       // //ABSOLUTE ENCODER
       IF #VTD_Control.AE_Error > 0 THEN
           "Set_Bit_F"(Bit := 5,
                       Bit_Value := 1,
                       Var := #VTD_Control.VTD_Errors.Error_Word_3);
       END_IF;

       //Errors while running
       IF #VTD_Control.Running THEN
           IF NOT (#VTD_Control.LP_State = 2) AND
               (#VTD_Control.LE > (#VTD_Settings.Teach_Values.Levels_LE[#LevelBelowExtractor] + #VTD_Settings.Slowdown_Count_LE) AND #VTD_Control.Instruction.Manual_Down)
               OR
               #IEC_Timer_0_Instance.Q
           THEN //22:4
               "Set_Bit_F"(Bit := 11,
                           Bit_Value := 1,
                           Var := #VTD_Control.VTD_Errors.Error_Word_1);
           END_IF;

           IF #VTD_Control.VFD_Error > 0 THEN //25:1
               "Set_Bit_F"(Bit := 0,
                           Bit_Value := 1,
                           Var := #VTD_Control.VTD_Errors.Error_Word_4);
           ELSIF #VTD_Control.LE_Error > 0 THEN //25:2
               "Set_Bit_F"(Bit := 1,
                           Bit_Value := 1,
                           Var := #VTD_Control.VTD_Errors.Error_Word_4);
           ELSIF #VTD_Control.AE_Error > 0 THEN //25:3
               "Set_Bit_F"(Bit := 2,
                           Bit_Value := 1,
                           Var := #VTD_Control.VTD_Errors.Error_Word_4);
           ELSIF (#LPL_Extended AND #LPL_Retracted) OR (#LPR_Extended AND #LPR_Retracted) THEN // 25:4
               "Set_Bit_F"(Bit := 3,
                           Bit_Value := 1,
                           Var := #VTD_Control.VTD_Errors.Error_Word_4);
           ELSIF #Lower_Limit AND NOT #Upper_limit THEN // 25:5
               "Set_Bit_F"(Bit := 4,
                           Bit_Value := 1,
                           Var := #VTD_Control.VTD_Errors.Error_Word_4);
           ELSIF NOT #Lower_Limit AND #Upper_limit THEN // 25:6
               "Set_Bit_F"(Bit := 5,
                           Bit_Value := 1,
                           Var := #VTD_Control.VTD_Errors.Error_Word_4);
           ELSIF #Lower_Limit AND #Upper_limit THEN // 25:7
               "Set_Bit_F"(Bit := 6,
                           Bit_Value := 1,
                           Var := #VTD_Control.VTD_Errors.Error_Word_4);
           END_IF;
       END_IF;

       //Check if overtravel limit switches has been hit
       IF #Upper_limit AND #Ultimate_Slow AND #Ulitmate_Creep AND #VTD_Control.Instruction.Manual_Up
       THEN //24:6 Top overtravel limit reached.
           "Set_Bit_F"(Bit := 7,
                       Bit_Value := 1,
                       Var := #VTD_Control.VTD_Errors.Error_Word_2);
           IF #VTD_Control.Mode = 2 OR #VTD_Control.Mode = 3 THEN
               #State := 400;
           ELSE
               #State := 0;
           END_IF;
       ELSIF #Lower_Limit AND #Ultimate_Slow AND #Ulitmate_Creep AND #VTD_Control.Instruction.Manual_Down
       THEN //24:7 Bottom overtravel limit reached.
               #VTD_Control.Error := TRUE; 
               "Set_Bit_F"(Bit := 8,
                           Bit_Value := 1,
                           Var := #VTD_Control.VTD_Errors.Error_Word_2);
               IF #VTD_Control.Mode = 2 OR #VTD_Control.Mode = 3 THEN
                   #State := 400;
               ELSE
                   #State := 0;
               END_IF;
       // ELSIF #Lower_Limit AND #Ultimate_Slow AND #Ulitmate_Creep AND #VTD_Control.Mode <> 4 THEN
       //     #VTD_Control.Instruction.Stop := TRUE;
       //     #VTD_Control.Error := TRUE; //24:7 Bottom Overtravel limit reached.
       //     "Set_Bit_F"(Bit := 8,
       //                 Bit_Value := 1,
       //                 Var := #VTD_Control.VTD_Errors.Error_Word_2);
       //     IF #VTD_Control.Mode = 2 OR #VTD_Control.Mode = 3 THEN
       //         #State := 400;
       //     ELSE
       //         #State := 0;
       //     END_IF;
       END_IF;

       //Need to monitor both encoders to (Need to uncomment)
       // #VTD_Control.Encoder_Delta := (#VTD_Control.LE - ((#VTD_Control.AE * #VTD_Settings.AE_Ratio)) * #VTD_Settings.Encoder_Delta_W1) + (#VTD_Control.Encoder_Delta * #VTD_Settings.Encoder_Delta_W2);
       IF ABS(#VTD_Control.Encoder_Delta) > #VTD_Settings.Encoder_Delta_Warning THEN
           //Send warning message that encoder error is to large
           #VTD_Control.Warning := 0;
       END_IF;

       "IEC_Timer_0_DB_10".TON(IN:=ABS(#VTD_Control.Encoder_Delta) > #VTD_Settings.Encoder_Delta_Error,
                               PT:=t#500ms);

       IF "IEC_Timer_0_DB_10".Q THEN
           //Send error message that encoder error is to large
           #VTD_Control.Error := TRUE; // 24:1
           "Set_Bit_F"(Bit := 2,
                       Bit_Value := 1,
                       Var := #VTD_Control.VTD_Errors.Error_Word_2);
           #State := 400;
       END_IF;

       // Level detect timer 
       IF #LD_Timer.Q THEN
           #LD_Timer(IN := FALSE,
                     PT := T#0s);
           #VTD_Control.Error := TRUE; // 24:10 VTD not level
           "Set_Bit_F"(Bit := 11,
                       Bit_Value := 1,
                       Var := #VTD_Control.VTD_Errors.Error_Word_4);
           #State := 400;
       END_IF;

       //Locking pin timer
       IF #LP_Timer.Q AND (#LPL_Retract OR #LPL_Extend) THEN //24:2 Locking pins took to long to extend
           "Set_Bit_F"(Bit := 3,
                       Bit_Value := 1,
                       Var := #VTD_Control.VTD_Errors.Error_Word_2);
       ELSIF #LP_Timer.Q AND (#LPR_Retract AND #LPR_Extend) THEN //24:3 Locking pins took to long to retract
           "Set_Bit_F"(Bit := 4,
                       Bit_Value := 1,
                       Var := #VTD_Control.VTD_Errors.Error_Word_2);
       END_IF;

       IF #Interlock_Timer.Q THEN //Interlock process timed out
           "Set_Bit_F"(Bit := 3,
                       Bit_Value := 1,
                       Var := #VTD_Control.VTD_Errors.Error_Word_3);
           #I_State := 400;
       END_IF;

       // Watchdog bit
       IF #Watchdog.Q THEN
           #VTD_Control.Running := FALSE;
           IF #VTD_Control.Mode = 4 THEN //24:9 Teach timed out
               "Set_Bit_F"(Bit := 10,
                           Bit_Value := 1,
                           Var := #VTD_Control.VTD_Errors.Error_Word_2);
           ELSIF #VTD_Control.Mode = 3 THEN //24:9 Auto timed out
               "Set_Bit_F"(Bit := 10,
                           Bit_Value := 1,
                           Var := #VTD_Control.VTD_Errors.Error_Word_2);
           ELSIF #VTD_Control.Mode = 2 THEN //24:9 Semi auto timed out
               "Set_Bit_F"(Bit := 10,
                           Bit_Value := 1,
                           Var := #VTD_Control.VTD_Errors.Error_Word_2);
           END_IF;
       END_IF;

       // go to error state
       IF  #VTD_Control.VTD_Errors.Error_Word_1 <> 0 OR
           #VTD_Control.VTD_Errors.Error_Word_2 <> 0 OR
           #VTD_Control.VTD_Errors.Error_Word_3 <> 0 OR
           #VTD_Control.VTD_Errors.Error_Word_4 <> 0 THEN
           #VTD_Control.Error := TRUE;
           #State := 400;
       END_IF;
   END_REGION

   REGION VFD
       //Status
       #VTD_Control.Motor.Ready := #SinaSpeed.Status = 16#7002;
       #VTD_Control.Motor.Running := #SinaSpeed.AxisEnabled;
       #VTD_Control.Motor.Error := #SinaSpeed.Status > 16#8000;

       //SETPOINT
       IF #VTD_Control.Motor_UP THEN
           #MainSetpoint := SCALE_X(MIN := 0,
                                    VALUE := NORM_X(MIN := 0,
                                                    VALUE := #VTD_Control.Motor_Speed,
                                                    MAX := 100),
                                    MAX := 1774);
       ELSIF #VTD_Control.Motor_Down THEN
           #MainSetpoint := (SCALE_X(MIN := 0,
                                     VALUE := NORM_X(MIN := 0,
                                                     VALUE := #VTD_Control.Motor_Speed,
                                                     MAX := 100),
                                     MAX := 1774)) * -1;
       ELSE
           #MainSetpoint := 0;
       END_IF;

       "IEC_Timer_0_DB".TON(IN:=#MainSetpoint <> 0,
                            PT:=T#500ms);

       IF "IEC_Timer_0_DB".Q THEN
           #MainSetpoint1 := #MainSetpoint;
       ELSE
           #MainSetpoint1 := 0;
       END_IF;

       IF #VTD_Control.Instruction.Enable THEN
           #SinaSpeed(EnableAxis := #VTD_Control.Motor_UP OR #VTD_Control.Motor_Down,
                          AckError := #VTD_Control.Instruction.Reset,
                          SpeedSp := #MainSetpoint1,
                          RefSpeed := 1774,
                          HWIDSTW := "VTD~PROFINET_interface~Standard_telegram_1",
                          HWIDZSW := "VTD~PROFINET_interface~Standard_telegram_1",
                          AxisEnabled => #VTD_Control.Motor.Status.%X0,
                          Lockout => #VTD_Control.Motor.Error,
                          Error => #VTD_Control.Motor.Error);
       END_IF;

       REGION Actual Speed
           IF #MainSetpoint1 > 0 THEN
               #VTD_Control.Motor.Speed_Actual := SCALE_X(MIN := 0,
                                                          VALUE := NORM_X(MIN := 0,
                                                                          VALUE := #SinaSpeed.ActVelocity,
                                                                          MAX := 1774),
                                                          MAX := 100);
           ELSIF #MainSetpoint1 < 0 THEN
               #VTD_Control.Motor.Speed_Actual := SCALE_X(MIN := 0,
                                                          VALUE := NORM_X(MIN := 0,
                                                                          VALUE := #SinaSpeed.ActVelocity * -1,
                                                                          MAX := 1774),
                                                          MAX := 100);
           ELSE
               #VTD_Control.Motor.Speed_Actual := 0;
           END_IF;
       END_REGION
   END_REGION

   //Assign local vars to outputs
   "Left LockingPin CMD Retract" := #LPL_Retract;
   "Left LockingPin CMD Extend" := #LPL_Extend;
   "Right LockingPin CMD Retract" := #LPR_Retract;
   "Right LockingPin CMD Extend" := #LPR_Extend;
END_FUNCTION_BLOCK

FUNCTION_BLOCK "EConveyor_FB"   // FB12, SCL
TITLE = Conveyor Instance FB
{ S7_Optimized_Access := 'TRUE' }
AUTHOR : Mertin Coetzee
VERSION : 0.1
// stored: AutoNumber true, IsIECCheckEnabled false, IsRetainMemResEnabled false, MemoryReserve 100, SetENOAutomatically false, UDAEnableTagReadback false
   VAR_INPUT
      Cnv_Settings : "ECnv_Settings";
      Cnv_Inputs : "ECnv_Inputs";
      VTD_Level : UInt;
      Cnv_TIP : Bool;
   END_VAR
   VAR_IN_OUT
      Cnv_Control : "ECnv_Control";
      SinaSpeed : SinaSpeed;
   END_VAR
   VAR
      State : UInt;
      Timer_TC : TON_TIME;
      Timer_Transfer { S7_SetPoint := 'True'} : TON_TIME;
      Watchdog { S7_SetPoint := 'True'} : TON_TIME;
      Transfer_Direction { S7_SetPoint := 'True'} : String;
      MainSetpoint : Int;
      SinaSpeed_Instance { S7_SetPoint := 'True'} : SinaSpeed;
      IEC_Timer_0_Instance_1 { S7_SetPoint := 'True'} : TON_TIME;
      IEC_Timer_0_Instance_2 { S7_SetPoint := 'True'} : TON_TIME;
      R_TRIG_Instance { S7_SetPoint := 'True'} : R_TRIG;
   END_VAR
   VAR_TEMP
      Execute_Old : Bool;
      Stop_Old : Bool;
      i : Int;
   END_VAR
BEGIN
   "R_TRIG_DB_15"(CLK := #Cnv_Control.Instruction.Execute AND NOT #Execute_Old);
   "R_TRIG_DB_16"(CLK := #Cnv_Control.Instruction.Stop AND NOT #Stop_Old);

   #Execute_Old := #Cnv_Control.Instruction.Execute;
   #Stop_Old := #Cnv_Control.Instruction.Stop;

   #Cnv_Control.Enabled := #Cnv_Control.Instruction.Enable;

   //MODES
   #Cnv_Control.Mode := #Cnv_Control.Instruction.Mode_Change;
   IF (#Cnv_Control.Mode = 1 OR #Cnv_Control.Mode = 5) AND NOT #Cnv_Control.Error THEN
       #State := 500;
   END_IF;

   #R_TRIG_Instance(CLK:=#Cnv_Control.Mode = 3);
   IF #R_TRIG_Instance.Q THEN
       #State := 0;
   END_IF;

   (*
   TODO:
   01. Need to add statemachine watchdog - Done
   02. Extractor needs to be on same floor for pallet to be moved in manual passed Rbwd - Done
   03. Complete reset state - Done
   04. Add stop inputs - Done
   05. Need to add variable motor speed, manual needs to be slower. - Done
   06. Need to add cyclic error checking. For odd sensor combinations as well - Partially done
   07. Need to add Shuttle monitor - Done
   08. Need to add Task ID check and start bit check to outbound pallet move. Check direction of pallet movement based on connected Cnv.
   09. Need to add checks for wrong direction of travel - Done
   10. Add checks for unsafe conditions with Cnv_Inputs - Partially Done
   11. Define Error codes - DOne
   12. Add watchdof time to Cnv Settings - Done
   13. Add self-timeout on manual 
   14. For shuttle in place sensor checks take into account extractor floor and safety stopper state
   15. Confirm modes and states are correct (Semi-auto and maintenance as well)
   16. Add the correct transfer process for the logistex-spacemaker pallet handovers.

   Mode select is done via the HMI. Might add external mode select switches.

           Mode select mask:
           0: Disabled
           1: Manual
           2: Semi-Auto
           3: Auto
           4: Teach - N/A for Cnv
           5: Maintenance

   Device ID Format: XXYYZZ    
   XX = Device type   
       01   VTD
       10  Cnv_Front_of_VTD
       11  Cnv_Rear_of_VTD
       12  Cnv_On_Extractor
       20  Safety_Stop_Front_of_VTD
       21  Safety_Stop_Rear_of_VTD
   YY = Floor   
   ZZ = VTD Connected to    
   Example: 110203 Conveyor at the rear of VTD 3 on level 2


    Sensor order for the conveyor:
    Lfwd Lpd1 Lpd2
     []   []   []
    ##############################
    #        Pallet Flow         #
    #         ------->>          #
    #                            #
    #                            #
    ##############################
                     []   []   []
                    Rpd2 Rpd1 Rbwd      
   *)

   REGION Cyclic Checks 
       #Cnv_Control.Cnv_Occupied := "Pallet in Position Rear VTD" AND "Pallet in Position Front VTD";

       //Check if a shuttle is in the Cnv
       FOR #i := 1 TO 3 DO
           IF "Shuttle_MQTT_DB".Shuttle_MQTT[#i].Message.Shuttle_Status.Position_ID = #Cnv_Settings.Barcode_ID THEN
               IF #Cnv_Inputs.Sdetect1 AND #Cnv_Inputs.Sdetect2 THEN
                   #Cnv_Control.Shuttle_In_Place := TRUE;
               ELSE
                   #Cnv_Control.Shuttle_In_Place := FALSE;
               END_IF;
           END_IF;
       END_FOR;

       // Update the Cnv_Control opbject
       #Cnv_Control.SM_State := #State;
       IF #Cnv_Control.Instruction.Inbound_Ready OR #Cnv_Control.Instruction.Outbound_Ready THEN
           #Cnv_Control.Ready_For_Task := TRUE;
       ELSE
           #Cnv_Control.Ready_For_Task := FALSE;
       END_IF;

   END_REGION

   REGION Auto/Semi/Manual mode
       CASE #State OF
           0: //IDLE MODE
               #Cnv_Control.Instruction.Transfer_Complete := 0;
               #Cnv_Control.Instruction.Transfer_in_Progress := FALSE;
               #Cnv_Control.Running := FALSE;
               #Cnv_Control.Motor.Forward := FALSE;
               #Cnv_Control.Motor.Reverse := FALSE;
               #Cnv_Control.Motor.Speed := 0;
               #Timer_Transfer(IN := FALSE,
                               PT := T#0S);
               IF #Cnv_Control.Enabled AND (#Cnv_Control.Mode = 3 OR #Cnv_Control.Mode = 2) AND #Cnv_Control.Error = 0 THEN
                   #State := 10;
               END_IF;

           10: //Standby - Conveyor ready to receive instruction
               IF ("R_TRIG_DB_15".Q OR #Cnv_Control.Instruction.Start_Transfer) AND "Control_DB".VTD_Control.Current_Level = #Cnv_Settings.Cnv_Level THEN
                   //Inbound Transfer
                   IF #Cnv_Control.Instruction.Inbound_Ready AND NOT #Cnv_Control.Running AND #Cnv_Control.Error = 0 AND
                       ("Control_DB".VTD_Control.Current_Level > 0 OR "Control_DB".PopUp_Cnv[2].Inputs."Lift Down")
                   THEN
                       #Cnv_Control.Done := FALSE;
                           #Cnv_Control.Running := TRUE;
                           #Cnv_Control.Instruction.Transfer_in_Progress := TRUE;
                           #Cnv_Control.Current_Task_ID := #Cnv_Control.Instruction.Task_ID;
                           #State := 20;

                       //Outbound Transfer    
                       ELSIF #Cnv_Control.Instruction.Outbound_Ready AND NOT #Cnv_Control.Running AND #Cnv_Control.Error = 0 AND
                           ("Control_DB".VTD_Control.Current_Level > 0 OR "Control_DB".PopUp_Cnv[2].Inputs."Lift Down")
                       THEN
                           #Cnv_Control.Done := FALSE;
                           #Cnv_Control.Running := TRUE;
                           #Cnv_Control.Instruction.Transfer_in_Progress := TRUE;
                           #Cnv_Control.Current_Task_ID := #Cnv_Control.Instruction.Task_ID;
                           #State := 30;
                   ELSE
                       #Cnv_Control.Warning := 1;// No task that can be started, yet start bit has been made true.
                   END_IF;
               ELSIF #Cnv_Control.Instruction.Start_Transfer AND "Control_DB".VTD_Control.Current_Level <> #Cnv_Settings.Cnv_Level THEN
                   //Extracot not at the correct level
                   "Set_Bit_F"(Bit := 2,
                               Bit_Value := 1,
                               Var := #Cnv_Control.Cnv_Errors.Error_Word_3);
               END_IF;

               //----------------------- Pallet Movement Inbound -----------------------
           20: // Running Roller FOWARD
               #Cnv_Control.Running := TRUE;
               #Cnv_Control.Motor.Forward := TRUE;
               #Cnv_Control.Motor.Speed := #Cnv_Settings.Full_Speed;
               #Transfer_Direction := 'Foward';

               IF "R_TRIG_DB_16".Q OR #Cnv_Control.Cnv_Occupied THEN
                   #Cnv_Control.Done := TRUE;
                   #Cnv_Control.Motor.Speed := 0;
                   #Cnv_Control.Motor.Forward := FALSE;
                   #Cnv_Control.Running := FALSE;
                   #State := 0;
               END_IF;

               //Monitor the transfer progress
               #Timer_Transfer(IN := TRUE,
                               PT := UINT_TO_TIME(#Cnv_Settings.Transfer_Time) * 1000);
               //If the watchdog bites, kill the process
               IF #Timer_Transfer.Q THEN //14:1 Transfer timed out
                   "Set_Bit_F"(Bit := 3,
                               Bit_Value := 1,
                               Var := #Cnv_Control.Cnv_Errors.Error_Word_2);
               END_IF;

               //----------------------- Pallet Movement Outbound -----------------------
           30: // Running Roller REVERSE
               IF (#VTD_Level = 0 AND "Control_DB".PopUp_Cnv[2].Chain_Motor.Status.%X0) OR
                   (#VTD_Level = 1 AND "Control_DB".LCnv_Control[1].Motor.Status.%X0) OR
                   (#VTD_Level = 2 AND "Control_DB".LCnv_Control[2].Motor.Status.%X0) OR
                   (#VTD_Level = 3 AND "Control_DB".LCnv_Control[3].Motor.Status.%X0) THEN
                   #Cnv_Control.Running := TRUE;
                   #Cnv_Control.Motor.Reverse := TRUE;
                   #Cnv_Control.Motor.Speed := #Cnv_Settings.Full_Speed;
                   #Transfer_Direction := 'Foward';
               END_IF;

               IF ("R_TRIG_DB_16".Q AND #Cnv_Control.Mode = 2) OR
                   (
                   (#VTD_Level = 0 AND NOT "PopUp Conveyor 2 - Pallet present 5") OR
                   (#VTD_Level = 1 AND NOT "Control_DB".LCnv_Control[1].Inputs."Pallet Detect 3") OR
                   (#VTD_Level = 2 AND NOT "Control_DB".LCnv_Control[2].Inputs."Pallet Detect 3") OR
                   (#VTD_Level = 3 AND NOT "Control_DB".LCnv_Control[3].Inputs."Pallet Detect 3") OR
                   (#VTD_Level = 99)
                   ) THEN
                   #Cnv_Control.Done := TRUE;
                   #Cnv_Control.Motor.Speed := 0;
                   #Cnv_Control.Motor.Forward := FALSE;
                   #Cnv_Control.Running := FALSE;
                   #State := 0;
               END_IF;

               //Monitor the transfer progress
               #Timer_Transfer(IN := TRUE,
                               PT := UINT_TO_TIME(#Cnv_Settings.Transfer_Time) * 1000);
               //If the watchdog bites, kill the process
               IF #Timer_Transfer.Q THEN //14:1 Transfer timed out
                   "Set_Bit_F"(Bit := 3,
                               Bit_Value := 1,
                               Var := #Cnv_Control.Cnv_Errors.Error_Word_2);
               END_IF;

           400: //Error state
               #Cnv_Control.Running := FALSE;
               #Cnv_Control.Motor.Speed := 0;
               #Cnv_Control.Motor.Forward := FALSE;
               #Cnv_Control.Motor.Reverse := FALSE;
               #Cnv_Control.Stopped := TRUE;
               #Cnv_Control.Instruction.Transfer_in_Progress := FALSE;
               #Watchdog(IN := FALSE,
                               PT := T#0S);
               #Timer_TC(IN := FALSE,
                               PT := T#0S);
               #Timer_Transfer(IN := FALSE,
                               PT := T#0S);
               #IEC_Timer_0_Instance_1(IN := FALSE,
                                       PT := T#0S);
               #IEC_Timer_0_Instance_2(IN := FALSE,
                                       PT := T#0S);
               IF #Cnv_Control.Instruction.Reset THEN
                   #Cnv_Control.Warning := 0;
                   #Cnv_Control.Current_Task_ID := 0;
                   #Cnv_Control.Error := FALSE; //Reset the conveyor

                   #Cnv_Control.Cnv_Errors.Error_Word_1 := 0;
                   #Cnv_Control.Cnv_Errors.Error_Word_2 := 0;
                   #Cnv_Control.Cnv_Errors.Error_Word_3 := 0;
                   #Cnv_Control.Cnv_Errors.Error_Word_4 := 0;
                   #State := 0;
               END_IF;

           500:
               IF #Cnv_Control.Enabled THEN
                   IF #"VTD_Level" = #Cnv_Settings.Cnv_Level THEN
                       IF #Cnv_Control.Instruction.Foward OR #Cnv_Control.Instruction.Start_Transfer THEN
                           #Cnv_Control.Motor.Speed := #Cnv_Settings.Manual_Speed;
                           #Cnv_Control.Motor.Forward := TRUE;
                           #Cnv_Control.Running := TRUE;
                       ELSIF #Cnv_Control.Instruction.Backward OR #Cnv_Control.Instruction.Start_Transfer_Backward THEN
                           #Cnv_Control.Motor.Speed := #Cnv_Settings.Manual_Speed;
                           #Cnv_Control.Motor.Reverse := TRUE;
                           #Cnv_Control.Running := TRUE;
                       ELSE
                           #Cnv_Control.Motor.Speed := 0;
                           #Cnv_Control.Motor.Forward := FALSE;
                           #Cnv_Control.Motor.Reverse := FALSE;
                           #Cnv_Control.Running := FALSE;
                       END_IF;
                   END_IF;
               END_IF;
               IF #Cnv_Control.Mode <> 1 AND #Cnv_Control.Mode <> 5 THEN
                   #State := 0;
               END_IF;
       END_CASE;
   END_REGION


   REGION Cyclic Error Checks
       IF NOT "Main_Safety_RTG1_DB".SAFETY_OK_VTD THEN //21:1
           "Set_Bit_F"(Bit := 0,
                       Bit_Value := 1,
                       Var := #Cnv_Control.Cnv_Errors.Error_Word_1);
       END_IF;

       IF #Cnv_Control.Motor.Error THEN
           "Set_Bit_F"(Bit := 0,
                       Bit_Value := 1,
                       Var := #Cnv_Control.Cnv_Errors.Error_Word_4);
       END_IF;


       // Shuttle in Place Cnv_Inputs - Need to confirm the order of these Cnv_Inputs.
       // IF (#Cnv_Settings.ID > 110000 AND #Cnv_Settings.ID < 120000 AND NOT #Cnv_Control.Inputs.Sdetect1 AND #Cnv_Control.Inputs.Sdetect2)
       //     OR (#Cnv_Settings.ID > 120000 AND #Cnv_Settings.ID < 130000 AND NOT #Cnv_Control.Inputs.Sdetect1 AND #Cnv_Control.Inputs.Sdetect2)
       // THEN //14:5 Shuttle is about to yeet itself down the VTD shaft
       //     "Set_Bit_F"(Bit := 7,
       //                 Bit_Value := 1,
       //                 Var := #Cnv_Control.Cnv_Errors.Error_Word_2);
       // END_IF;

       // IF (#Cnv_Settings.ID > 110000 AND #Cnv_Settings.ID < 120000 AND #Cnv_Control.Inputs.Sdetect1 AND NOT #Cnv_Control.Inputs.Sdetect2)
       //     OR (#Cnv_Settings.ID > 120000 AND #Cnv_Settings.ID < 130000 AND #Cnv_Control.Inputs.Sdetect1 AND NOT #Cnv_Control.Inputs.Sdetect2) THEN
       //     #Cnv_Control.Warning := 1; //Shuttle detected in conveyor not yet on barcode
       // END_IF;

       //Watchdog auto starts the moment any form of transfer occurs.
       // IF #State > 10 AND #State < 400 THEN
       //     #Watchdog(IN := TRUE,
       //               PT := T#600s);
       // ELSE
       //     #Watchdog.IN := FALSE;
       // END_IF;

       // IF #Watchdog.Q THEN
       //     #Watchdog.IN := FALSE;
       //     #Cnv_Control.Error := TRUE; //14:2  Watchdog bit
       //     "Set_Bit_F"(Bit := 4,
       //                 Bit_Value := 1,
       //                 Var := #Cnv_Control.Cnv_Errors.Error_Word_2);
       //     #State := 400;
       // END_IF;

       // go to error state
       IF #Cnv_Control.Cnv_Errors.Error_Word_1 <> 0 OR
           #Cnv_Control.Cnv_Errors.Error_Word_2 <> 0 OR
           #Cnv_Control.Cnv_Errors.Error_Word_3 <> 0 OR
           #Cnv_Control.Cnv_Errors.Error_Word_4 <> 0
           THEN
               #Cnv_Control.Error := TRUE;
               #State := 400;
       END_IF;
   END_REGION

   REGION VFD
       //Status
       #Cnv_Control.Motor.Ready := NOT #Cnv_Control.Motor.Error;

       #SinaSpeed(EnableAxis := #Cnv_Control.Motor.Forward OR #Cnv_Control.Motor.Reverse,
                  AckError := #Cnv_Control.Instruction.Reset,
                  SpeedSp := #MainSetpoint,
                  RefSpeed := 1745.0,
                  HWIDSTW := #Cnv_Settings.G120_Hardware_ID,
                  HWIDZSW := #Cnv_Settings.G120_Hardware_ID,
                  AxisEnabled => #Cnv_Control.Motor.Status.%X0,
                  Lockout => #Cnv_Control.Motor.Error,
                  Error => #Cnv_Control.Motor.Error);

       //MAIN SETPOINT
       IF #Cnv_Control.Motor.Reverse THEN
           #MainSetpoint := (SCALE_X(MIN := 0,
                                    VALUE := NORM_X(MIN := 0,
                                                    VALUE := #Cnv_Control.Motor.Speed,
                                                    MAX := 100),
                                    MAX := 1745.0)) * -1;
      ELSIF #Cnv_Control.Motor.Forward THEN
           #MainSetpoint := SCALE_X(MIN := 0,
                                     VALUE := NORM_X(MIN := 0,
                                                     VALUE := #Cnv_Control.Motor.Speed,
                                                     MAX := 100),
                                     MAX := 1745.0);
       ELSE
           #MainSetpoint := 0;
       END_IF;

       //Actual Speed
       IF #MainSetpoint > 0 THEN
           #Cnv_Control.Motor.Speed_Actual := SCALE_X(MIN := 0,
                                                      VALUE := NORM_X(MIN := 0,
                                                                      VALUE := #SinaSpeed.ActVelocity,
                                                                      MAX := 1745.0),
                                                      MAX := 100);
       ELSIF #MainSetpoint < 0 THEN
           #Cnv_Control.Motor.Speed_Actual := SCALE_X(MIN := 0,
                                                      VALUE := NORM_X(MIN := 0,
                                                                      VALUE := #SinaSpeed.ActVelocity * -1,
                                                                      MAX := 1745.0),
                                                      MAX := 100);
       ELSE
           #Cnv_Control.Motor.Speed_Actual := 0;
       END_IF;
   END_REGION
END_FUNCTION_BLOCK

FUNCTION_BLOCK "Buffer_Conveyor_FB"   // FB5, SCL
TITLE = Conveyor Instance FB
{ S7_Optimized_Access := 'TRUE' }
AUTHOR : Mertin Coetzee
VERSION : 0.1
// stored: AutoNumber true, IsIECCheckEnabled false, IsRetainMemResEnabled false, MemoryReserve 100, SetENOAutomatically false, UDAEnableTagReadback false
   VAR_INPUT
      Cnv_Settings : "Buffer_Cnv_Settings";
      VTD_Level : UInt;
      ECnv_TIP : Bool;
   END_VAR
   VAR_IN_OUT
      Cnv_Control : "Buffer_Cnv_Control";
      SinaSpeed : SinaSpeed;
   END_VAR
   VAR
      State : UInt;
      Timer_TC : TON_TIME;
      Timer_Transfer { S7_SetPoint := 'True'} : TON_TIME;
      Watchdog { S7_SetPoint := 'True'} : TON_TIME;
      Transfer_Direction { S7_SetPoint := 'True'} : String;
      MainSetpoint : Int;
      IEC_Timer_0_Instance_1 { S7_SetPoint := 'True'} : TON_TIME;
      R_TRIG_Instance { S7_SetPoint := 'True'} : R_TRIG;
   END_VAR
   VAR_TEMP
      Execute_Old : Bool;
      Stop_Old : Bool;
   END_VAR
BEGIN
   "R_TRIG_DB_17"(CLK := #Cnv_Control.Instruction.Execute AND NOT #Execute_Old);
   "R_TRIG_DB_18"(CLK := #Cnv_Control.Instruction.Stop AND NOT #Stop_Old);

   #Execute_Old := #Cnv_Control.Instruction.Execute;
   #Stop_Old := #Cnv_Control.Instruction.Stop;

   #Cnv_Control.Enabled := #Cnv_Control.Instruction.Enable;

   //MODES
   #Cnv_Control.Mode := #Cnv_Control.Instruction.Mode_Change;
   IF (#Cnv_Control.Mode = 1 OR #Cnv_Control.Mode = 5) AND NOT #Cnv_Control.Error THEN
       #State := 500;
   END_IF;

   #R_TRIG_Instance(CLK:=#Cnv_Control.Mode = 3);
   IF #R_TRIG_Instance.Q THEN
       #State := 0;
   END_IF;

   (*
   TODO:
   01. Need to add statemachine watchdog - Done
   02. Extractor needs to be on same floor for pallet to be moved in manual passed Rbwd - Done
   03. Complete reset state - Done
   04. Add stop inputs - Done
   05. Need to add variable motor speed, manual needs to be slower. - Done
   06. Need to add cyclic error checking. For odd sensor combinations as well - Partially done
   07. Need to add Shuttle monitor - Done
   08. Need to add Task ID check and start bit check to outbound pallet move. Check direction of pallet movement based on connected Cnv.
   09. Need to add checks for wrong direction of travel - Done
   10. Add checks for unsafe conditions with Cnv_Inputs - Partially Done
   11. Define Error codes - DOne
   12. Add watchdof time to Cnv Settings - Done
   13. Add self-timeout on manual 
   14. For shuttle in place sensor checks take into account extractor floor and safety stopper state
   15. Confirm modes and states are correct (Semi-auto and maintenance as well)
   16. Add the correct transfer process for the logistex-spacemaker pallet handovers.

   Mode select is done via the HMI. Might add external mode select switches.

           Mode select mask:
           0: Disabled
           1: Manual
           2: Semi-Auto
           3: Auto
           4: Teach - N/A for Cnv
           5: Maintenance

   Device ID Format: XXYYZZ    
   XX = Device type   
       40  VTD
       10  Cnv_Front_of_VTD
       11  Cnv_Rear_of_VTD
       12  Cnv_On_Extractor
       20  Safety_Stop_Front_of_VTD
       21  Safety_Stop_Rear_of_VTD

   YY = Floor   
   ZZ = VTD Connected to    
   Example: 110203 Conveyor at the rear of VTD 3 on level 2

   Pallet Alignment
   0 = no alignment
   1 = center alignment
   2 = Left
   3 = Right

    Sensor order for the conveyor:
    Lfwd Lpd1 Lpd2
     []   []   []
    ##############################
    #        Pallet Flow         #
    #         ------->>          #
    #                            #
    #                            #
    ##############################
                     []   []   []
                    Rpd2 Rpd1 Rbwd      
   *)

   REGION Cyclic Checks    
       #Cnv_Control.Cnv_Occupied := NOT #Cnv_Control.Inputs."Pallet Detect 1" AND (*#Cnv_Control."Inputs"."Pallet Detect 2" AND*) NOT #Cnv_Control.Inputs."Pallet Detect 3";

       //Check if a shuttle is in the Cnv
       IF NOT #Cnv_Control.Inputs.Sdetect1 AND NOT #Cnv_Control.Inputs.Sdetect2 THEN
           #Cnv_Control.Shuttle_In_Place := TRUE;
       ELSE
           #Cnv_Control.Shuttle_In_Place := FALSE;
       END_IF;

       // Update the Cnv_Control opbject
       #Cnv_Control.SM_State := #State;
       #Cnv_Control.Stopped := NOT #Cnv_Control.Running;
       IF #Cnv_Control.Instruction.Inbound_Ready OR #Cnv_Control.Instruction.Outbound_Ready THEN
           #Cnv_Control.Ready_For_Task := TRUE;
       ELSE
           #Cnv_Control.Ready_For_Task := FALSE;
       END_IF;

   END_REGION

   REGION Auto/Semi auto mode
       CASE #State OF
           0: //Initialization
               #Cnv_Control.Instruction.Transfer_Complete := 0;
               #Cnv_Control.Instruction.Transfer_in_Progress := FALSE;
               #Cnv_Control.Running := FALSE;
               #Cnv_Control.Motor.Forward := FALSE;
               #Cnv_Control.Motor.Reverse := FALSE;
               #Cnv_Control.Motor.Speed := 0;
               #Timer_Transfer(IN := FALSE,
                               PT := T#0S);
               IF #Cnv_Control.Enabled AND (#Cnv_Control.Mode = 3 OR #Cnv_Control.Mode = 2) AND #Cnv_Control.Error = 0 THEN
                   #State := 10;
               END_IF;

               10: //Standby - Conveyor ready to receive instruction
                   IF ("R_TRIG_DB_17".Q OR #Cnv_Control.Instruction.Start_Transfer) AND "Control_DB".VTD_Control.Current_Level = #Cnv_Settings.Cnv_Level THEN
                       //Inbound Transfer
                       IF #Cnv_Control.Instruction.Inbound_Ready AND NOT #Cnv_Control.Running AND #Cnv_Control.Error = 0 THEN
                           //Check transfer ID
                           #Cnv_Control.Done := FALSE;
                               #Cnv_Control.Running := TRUE;
                               #Cnv_Control.Instruction.Transfer_in_Progress := TRUE;
                               #Cnv_Control.Current_Task_ID := #Cnv_Control.Instruction.Task_ID;
                               #State := 20;

                           //Outbound Transfer    
                       ELSIF #Cnv_Control.Instruction.Outbound_Ready AND NOT #Cnv_Control.Running AND #Cnv_Control.Error = 0 THEN
                           //Check transfer ID
                           #Cnv_Control.Done := FALSE;
                               #Cnv_Control.Running := TRUE;
                               #Cnv_Control.Instruction.Transfer_in_Progress := TRUE;
                               #Cnv_Control.Current_Task_ID := #Cnv_Control.Instruction.Task_ID;
                               #State := 30;
                       ELSE
                           #Cnv_Control.Warning := 0;// No task that can be started, yet start bit has been made true.
                       END_IF;
                   ELSIF #Cnv_Control.Instruction.Start_Transfer AND "Control_DB".VTD_Control.Current_Level <> #Cnv_Settings.Cnv_Level THEN
                       //Extractor not at the correct level
                       "Set_Bit_F"(Bit := 2,
                                   Bit_Value := 1,
                                   Var := #Cnv_Control.Cnv_Errors.Error_Word_3);
                   END_IF;

                   //----------------------- Pallet Movement Inbound -----------------------
               20: // Running Roller FOWARD
                   #Cnv_Control.Running := TRUE;
                   #Cnv_Control.Motor.Forward := TRUE;
                   #Cnv_Control.Motor.Speed := #Cnv_Settings.Full_Speed;
                   #Transfer_Direction := 'Foward';

                   IF "R_TRIG_DB_18".Q OR NOT #Cnv_Control.Inputs."Pallet Detect 3" THEN
                       #Cnv_Control.Done := TRUE;
                       #Cnv_Control.Motor.Speed := 0;
                       #Cnv_Control.Motor.Forward := FALSE;
                       #Cnv_Control.Running := FALSE;
                       #State := 0;
                   END_IF;

                   //Monitor the transfer progress
                   #Timer_Transfer(IN := TRUE,
                                   PT := UINT_TO_TIME(#Cnv_Settings.Transfer_Time) * 1000);
                   //If the watchdog bites, kill the process
                   IF #Timer_Transfer.Q THEN //14:1 Transfer timed out
                       "Set_Bit_F"(Bit := 3,
                                   Bit_Value := 1,
                                   Var := #Cnv_Control.Cnv_Errors.Error_Word_2);
                   END_IF;

                   //----------------------- Pallet Movement Outbound -----------------------
               30: // Running Roller REVERSE
                   #Cnv_Control.Running := TRUE;
                   #Cnv_Control.Motor.Reverse := TRUE;
                   #Cnv_Control.Motor.Speed := #Cnv_Settings.Full_Speed;
                   #Transfer_Direction := 'Foward';

                   IF "R_TRIG_DB_18".Q OR "Control_DB".ECnv_Control.Cnv_Occupied THEN
                       #Cnv_Control.Done := TRUE;
                       #Cnv_Control.Motor.Speed := 0;
                       #Cnv_Control.Motor.Forward := FALSE;
                       #Cnv_Control.Running := FALSE;
                       #State := 0;
                   END_IF;

                   //Monitor the transfer progress
                   #Timer_Transfer(IN := TRUE,
                                   PT := UINT_TO_TIME(#Cnv_Settings.Transfer_Time) * 1000);
                   //If the watchdog bites, kill the process
                   IF #Timer_Transfer.Q THEN //14:1 Transfer timed out
                       "Set_Bit_F"(Bit := 3,
                                   Bit_Value := 1,
                                   Var := #Cnv_Control.Cnv_Errors.Error_Word_2);
                   END_IF;

               400: //Error state
                   #Cnv_Control.Running := FALSE;
                   #Cnv_Control.Motor.Speed := 0;
                   #Cnv_Control.Motor.Forward := FALSE;
                   #Cnv_Control.Motor.Reverse := FALSE;
                   #Cnv_Control.Instruction.Stop := FALSE;
                   #Cnv_Control.Instruction.Transfer_in_Progress := FALSE;
                   #Watchdog(IN := FALSE,
                                   PT := T#0S);
                   #Timer_TC(IN := FALSE,
                                   PT := T#0S);
                   #Timer_Transfer(IN := FALSE,
                                   PT := T#0S);
                   #IEC_Timer_0_Instance_1(IN := FALSE,
                                           PT := T#0S);
                   IF #Cnv_Control.Instruction.Reset THEN
                       #Cnv_Control.Warning := 0;
                       #Cnv_Control.Current_Task_ID := 0;
                       #Cnv_Control.Error := FALSE; //Reset the conveyor

                       #Cnv_Control.Cnv_Errors.Error_Word_1 := 0;
                       #Cnv_Control.Cnv_Errors.Error_Word_2 := 0;
                       #Cnv_Control.Cnv_Errors.Error_Word_3 := 0;
                       #Cnv_Control.Cnv_Errors.Error_Word_4 := 0;
                       #State := 0;
                   END_IF;

               500:
                   IF #Cnv_Control.Enabled THEN
                       IF #Cnv_Control.Instruction.Foward OR #Cnv_Control.Instruction.Start_Transfer THEN
                               #Cnv_Control.Motor.Speed := #Cnv_Settings.Manual_Speed;
                               #Cnv_Control.Motor.Forward := TRUE;
                               #Cnv_Control.Running := TRUE;
                           ELSIF #Cnv_Control.Instruction.Backward OR #Cnv_Control.Instruction.Start_Transfer_Backward THEN
                               #Cnv_Control.Motor.Speed := #Cnv_Settings.Manual_Speed;
                               #Cnv_Control.Motor.Reverse := TRUE;
                               #Cnv_Control.Running := TRUE;
                           ELSE
                               #Cnv_Control.Motor.Speed := 0;
                               #Cnv_Control.Motor.Forward := FALSE;
                               #Cnv_Control.Motor.Reverse := FALSE;
                               #Cnv_Control.Running := FALSE;
                           END_IF;
                       END_IF;
                   IF #Cnv_Control.Mode <> 1 AND #Cnv_Control.Mode <> 5 THEN
                       #State := 0;
                   END_IF;
           END_CASE;
       END_REGION



   REGION Cyclic Error Checks
       IF NOT "Main_Safety_RTG1_DB".SAFETY_OK_VTD THEN //11:1
           "Set_Bit_F"(Bit := 0,
                       Bit_Value := 1,
                       Var := #Cnv_Control.Cnv_Errors.Error_Word_1);
       END_IF;

       // IF #Cnv_Control.Instruction.Stop THEN //11:2
       //     "Set_Bit_F"(Bit := 1,
       //                 Bit_Value := 1,
       //                 Var := #Cnv_Control.Cnv_Errors.Error_Word_1);
       // END_IF;

       IF #Cnv_Control.Motor.Error THEN
           "Set_Bit_F"(Bit := 0,
                       Bit_Value := 1,
                       Var := #Cnv_Control.Cnv_Errors.Error_Word_4);
       END_IF;

       // Pallet Sensor Checks
       // IF #Cnv_Control.Inputs.Lfwd AND #Cnv_Control.Inputs.Rbwd THEN
       //     #Cnv_Control.Error := TRUE; //15:2 Combination of Cnv_Inputs indicates issue in conveyor
       //     "Set_Bit_F"(Bit := 1,
       //                 Bit_Value := 1,
       //                 Var := #Cnv_Control.Cnv_Errors.Error_Word_4);
       //     #State := 400;
       // IF #Cnv_Control.Inputs.Lfwd AND #Cnv_Control.Inputs.Lpd1 AND #Cnv_Control.Inputs.Rpd1 THEN
       //     #Cnv_Control.Error := TRUE; //15:3 Combination of Cnv_Inputs indicates issue in conveyor
       //     "Set_Bit_F"(Bit := 2,
       //                 Bit_Value := 1,
       //                 Var := #Cnv_Control.Cnv_Errors.Error_Word_4);
       //     #State := 400;
       // ELSIF #Cnv_Control.Inputs.Rbwd AND #Cnv_Control.Inputs.Lpd1 AND #Cnv_Control.Inputs.Rpd1 THEN
       //     #Cnv_Control.Error := TRUE; //15:4 Combination of Cnv_Inputs indicates issue in conveyor
       //     "Set_Bit_F"(Bit := 3,
       //                 Bit_Value := 1,
       //                 Var := #Cnv_Control.Cnv_Errors.Error_Word_4);
       //     #State := 400;
       // END_IF;

       // Shuttle in Place Cnv_Inputs - Need to confirm the order of these Cnv_Inputs.
       // IF (#Cnv_Settings.ID > 110000 AND #Cnv_Settings.ID < 120000 AND NOT #Cnv_Control.Inputs.Sdetect1 AND #Cnv_Control.Inputs.Sdetect2)
       //     OR (#Cnv_Settings.ID > 120000 AND #Cnv_Settings.ID < 130000 AND NOT #Cnv_Control.Inputs.Sdetect1 AND #Cnv_Control.Inputs.Sdetect2) THEN
       //     #Cnv_Control.Error := TRUE; //14:5 Shuttle is about to yeet itself down the VTD shaft
       //     "Set_Bit_F"(Bit := 7,
       //                 Bit_Value := 1,
       //                 Var := #Cnv_Control.Cnv_Errors.Error_Word_2);
       //     #State := 400;
       // END_IF;

       // IF (#Cnv_Settings.ID > 110000 AND #Cnv_Settings.ID < 120000 AND #Cnv_Control.Inputs.Sdetect1 AND NOT #Cnv_Control.Inputs.Sdetect2)
       //     OR (#Cnv_Settings.ID > 120000 AND #Cnv_Settings.ID < 130000 AND #Cnv_Control.Inputs.Sdetect1 AND NOT #Cnv_Control.Inputs.Sdetect2) THEN
       //     #Cnv_Control.Warning := 0; //Shuttle detected in conveyor not yet on barcode
       // END_IF;

       // // #Watchdog auto starts the moment Any form OF transfer occurs.
       // IF #State > 10 AND #State < 400 THEN
       //     #Watchdog(IN := TRUE,
       //               PT := T#200s);
       // ELSE
       //     #Watchdog.IN := FALSE;
       // END_IF;

       // IF #Watchdog.Q THEN
       //     #Watchdog.IN := FALSE;
       //     #Cnv_Control.Error := TRUE; //14:2  Watchdog bit
       //     "Set_Bit_F"(Bit := 4,
       //                 Bit_Value := 1,
       //                 Var := #Cnv_Control.Cnv_Errors.Error_Word_2);
       //     #State := 400;
       // END_IF;

       // go to error state
       IF #Cnv_Control.Cnv_Errors.Error_Word_1 <> 0 OR
           #Cnv_Control.Cnv_Errors.Error_Word_2 <> 0 OR
           #Cnv_Control.Cnv_Errors.Error_Word_3 <> 0 OR
           #Cnv_Control.Cnv_Errors.Error_Word_4 <> 0
           THEN
               #Cnv_Control.Error := TRUE;
               #State := 400;
       END_IF;
   END_REGION

   REGION VFD
       //Status
       #Cnv_Control.Motor.Ready := NOT #Cnv_Control.Motor.Error;

       #SinaSpeed(EnableAxis := #Cnv_Control.Motor.Forward OR #Cnv_Control.Motor.Reverse,
                  AckError := #Cnv_Control.Instruction.Reset,
                  SpeedSp := #MainSetpoint,
                  RefSpeed := 1745.0,
                  HWIDSTW := #Cnv_Settings.G120_Hardware_ID,
                  HWIDZSW := #Cnv_Settings.G120_Hardware_ID,
                  AxisEnabled => #Cnv_Control.Motor.Status.%X0,
                  Lockout => #Cnv_Control.Motor.Error,
                  Error => #Cnv_Control.Motor.Error);

       //MAIN SETPOINT
       IF #Cnv_Control.Motor.Forward THEN
           #MainSetpoint := (SCALE_X(MIN := 0,
                                    VALUE := NORM_X(MIN := 0,
                                                    VALUE := #Cnv_Control.Motor.Speed * 1.681,
                                                    MAX := 100),
                                    MAX := 1745.0) * -1);
       ELSIF #Cnv_Control.Motor.Reverse THEN
           #MainSetpoint := SCALE_X(MIN := 0,
                                     VALUE := NORM_X(MIN := 0,
                                                     VALUE := #Cnv_Control.Motor.Speed * 1.681,
                                                     MAX := 100),
                                     MAX := 1745.0);
       ELSE
           #MainSetpoint := 0;
       END_IF;

       REGION Actual Speed
           IF #MainSetpoint > 0 THEN
               #Cnv_Control.Motor.Speed_Actual := SCALE_X(MIN := 0,
                                                          VALUE := NORM_X(MIN := 0,
                                                                          VALUE := #SinaSpeed.ActVelocity,
                                                                          MAX := 1745.0),
                                                          MAX := 100);
           ELSIF #MainSetpoint < 0 THEN
               #Cnv_Control.Motor.Speed_Actual := SCALE_X(MIN := 0,
                                                          VALUE := NORM_X(MIN := 0,
                                                                          VALUE := #SinaSpeed.ActVelocity * -1,
                                                                          MAX := 1745.0),
                                                          MAX := 100);
           ELSE
               #Cnv_Control.Motor.Speed_Actual := 0;
           END_IF;
       END_REGION
   END_REGION
END_FUNCTION_BLOCK

FUNCTION_BLOCK "Safety_Stops_FB"   // FB7, SCL
{ S7_Optimized_Access := 'TRUE' }
VERSION : 0.1
// stored: AutoNumber true, IsIECCheckEnabled false, IsRetainMemResEnabled false, MemoryReserve 100, SetENOAutomatically false, UDAEnableTagReadback false
   VAR_INPUT
      Mode : UInt;
      Timeout : UInt;
      Reset : Bool;
      Up : Bool;
      Down : Bool;
   END_VAR
   VAR_OUTPUT
      Rotate : Bool;
   END_VAR
   VAR_IN_OUT
      Sfts_Control : "Sfts_Control";
   END_VAR
   VAR
      State : UInt;
      LP_Timer { ExternalAccessible := 'False'; ExternalVisible := 'False'; ExternalWritable := 'False'} : TON_TIME;
      IEC_Timer_0_Instance { S7_SetPoint := 'True'} : TOF_TIME;
      Timer_1 : Time;
   END_VAR
BEGIN
   #Sfts_Control.Enabled := #Sfts_Control.Instruction.Enable := #Mode = 2 OR #Mode = 3;

   //MODES
   IF (#Mode = 1 OR #Mode = 5) AND NOT #Sfts_Control.Error THEN
       #State := 500;
   END_IF;

   (*
   TODO
   1. Need to add the mode and running checks for manual mode
   2. Add output for safety stop brake.

   Mode select is done via the HMI. Might add external mode select switches.

           Mode select mask:
           0: Disabled
           1: Manual
           2: Semi-Auto
           3: Auto
           4: Teach - N/A for Cnv
           5: Maintenance

   Device ID Format: XXYYZZ    
   XX = Device type   
       01   VTD
       10  Cnv_Front_of_VTD
       11  Cnv_Rear_of_VTD
       12  Cnv_On_Extractor
       20  Safety_Stop_Front_of_VTD
       21  Safety_Stop_Rear_of_VTD
   YY = Floor   
   ZZ = VTD Connected to 
   *)

   REGION Assign Inputs
       #Sfts_Control.Inputs.LP_Extended := #Up;
       #Sfts_Control.Inputs.LP_Retracted := #Down;
   END_REGION

   REGION Cyclic Checks
       //Update variables
       #Sfts_Control.SM_State := #State;

       #LP_Timer(IN := #Sfts_Control.Running,
                 PT := UINT_TO_TIME(#Timeout));

       //STOPPER STATE
       IF #Sfts_Control.Inputs.LP_Extended AND NOT #Sfts_Control.Inputs.LP_Retracted THEN
           #Sfts_Control.LP_State := 1; // EXTENDED
       ELSIF NOT #Sfts_Control.Inputs.LP_Extended AND #Sfts_Control.Inputs.LP_Retracted THEN
           #Sfts_Control.LP_State := 0; //RETRACTED
       ELSE
           #Sfts_Control.LP_State := 2; //LOST
       END_IF;;
   END_REGION

   REGION Auto Mode

           CASE #State OF
               0: //IDLE MODE
                   IF #Mode = 2 OR #Mode = 3 THEN
                       IF #Sfts_Control.Instruction.Enable AND #Sfts_Control.Error = 0 THEN
                           #Sfts_Control.Enabled := TRUE;
                           #State := 10;
                       END_IF;
                   END_IF;
               10: //Standby
                   IF NOT #Sfts_Control.Running AND #Sfts_Control.Error = 0 AND #Sfts_Control.Instruction.LP_Extend THEN
                       IF #Sfts_Control.Inputs.LP_Extended THEN
                           ; // Complete the task as the LP ar already extended
                       ELSIF #Sfts_Control.Inputs.LP_Retracted THEN
                           #Sfts_Control.Running := True;
                           #State := 20;
                       ELSE
                           #Sfts_Control.Error := 0; //Unknown locking pin state
                           #State := 400;
                       END_IF;
                   ELSIF NOT #Sfts_Control.Running AND #Sfts_Control.Error = 0 AND #Sfts_Control.Instruction.LP_Retract THEN
                       IF #Sfts_Control.Inputs.LP_Retracted THEN
                           ; // Complete the task as the LP ar already extended
                       ELSIF #Sfts_Control.Inputs.LP_Extended THEN
                           #Sfts_Control.Running := True;
                           #State := 40;
                       ELSE
                           #Sfts_Control.Error := 0; //Unknown locking pin state
                           #State := 400;
                       END_IF;
                   END_IF;

               20: //Extend safety locking pins
                   #Sfts_Control.Motor_Extend := TRUE;
                   IF #Sfts_Control.Inputs.LP_Extended THEN
                       #Sfts_Control.Motor_Extend := FALSE;
                       #Sfts_Control.Running := FALSE;
                       #State := 0;
                   END_IF;

               40: //Retract safety locking pins
                   #Sfts_Control.Motor_Retract := TRUE;
                   IF #Sfts_Control.Inputs.LP_Retracted THEN
                       #Sfts_Control.Motor_Retract := FALSE;
                       #Sfts_Control.Running := FALSE;
                       #State := 0;
                   END_IF;

               400: // Error#Sfts_Control
                   #Sfts_Control.Motor_Retract := FALSE;
                   #Sfts_Control.Motor_Extend := FALSE;
                   #Sfts_Control.Running := FALSE;
                   #LP_Timer(IN := FALSE,
                             PT := T#0S);
                   IF #Reset THEN
                       #Sfts_Control.Error := FALSE;
                       #State := 0;
                   END_IF;

               500:
                   IF #Sfts_Control.Instruction.Manual_Extend AND NOT #Sfts_Control.Inputs.LP_Extended THEN
                       #Sfts_Control.Motor_Extend := TRUE;
                       #Sfts_Control.Running := TRUE;
                   ELSIF #Sfts_Control.Instruction.Manual_Retract AND NOT #Sfts_Control.Inputs.LP_Retracted THEN
                       #Sfts_Control.Motor_Retract := TRUE;
                       #Sfts_Control.Running := TRUE;
                   ELSE
                       #Sfts_Control.Motor_Extend := FALSE;
                       #Sfts_Control.Motor_Retract := FALSE;
                       #Sfts_Control.Running := FALSE;
                   END_IF;

                   IF #Mode <> 1 AND #Mode <> 5 THEN
                       #State := 0;
                   END_IF;
           END_CASE;
   END_REGION

   REGION Cyclic Error Checks
       IF #Sfts_Control.Inputs.LP_Extended AND #Sfts_Control.Inputs.LP_Retracted THEN
           #Sfts_Control.Error := TRUE; //Cant have the locking pins extended and retracted at the same time11
       END_IF;

       // Statement section REGION
       IF #LP_Timer.Q THEN
           #Sfts_Control.Error := TRUE;//locking pin timeout
       END_IF;

       IF #Sfts_Control.Error THEN
           #State := 400;
       END_IF;
   END_REGION

   REGION Assign outputs
       #IEC_Timer_0_Instance(IN := #Sfts_Control.Motor_Extend OR #Sfts_Control.Motor_Retract,
                             PT := #Timer_1,
                             Q => #Rotate);
   END_REGION
END_FUNCTION_BLOCK

FUNCTION "Encoders" : Void   // FC8, SCL
{ S7_Optimized_Access := 'TRUE' }
VERSION : 0.1
// stored: AutoNumber true, IsIECCheckEnabled false, SetENOAutomatically false, UDAEnableTagReadback false
BEGIN
   REGION ABSOLUTE ENCODER
       //STATUS---------------------------------------------------------------------------------------------------------------------
       //
       //Encoder state word 2 - INPUT WORD 1
       //
       // 15 … 12 Encoder’s Sign-OF-Life (NOT relevant)
       // 11, 10 Reserved
       // 9 Control requested 0 = No control BY the PLC requested 1 = Control BY the PLC requested
       // 8 … 0 Reserved

       //Sensor 1 state word - INPUT WORD 2
       //
       // 15 Encoder error Description 0 = No error 1 = Error The error code is output in G1_XIST2.
       // 14 Park mode activated 0 = Normal operation 1 = Park mode activated Feedback based on G1_STW bit 14: No output OF position data G1_XIST1 AND G1_XIST2
       // 13 Transmission OF absolute position value 0 = No transmission 1 = Position value is output in G1_XIST2
       // 12 Status OF the Preset function (set/shift OF home position executed) 0 = No Preset function active 1 = Preset function is run Feedback based on G1_STW bit 12:  
       // 11 Requirement OF error acknowledgement detected New position value is output in G1_XIST1 AND G1_XIST2. On conclusion OF the Preset function the bit is set TO 0. 0 = No RETURN acknowledgement OF Encoder error 1 = Requirement OF error acknowledgement detected Reaction TO bit 15 in the sensor control word 1 G1_STW is acknowledged (see Table 14)
       // 10 Reserved
       // 9 … 0 NOT supported

       //Position 1 - INPUT WORD 3 AND 4
       // "AE_Position_1_Scaled" := (*SCALE_X(MIN := "Settings_DB".VTD_Settings.VTD_Min_Height,
       //                                   VALUE := *)NORM_X(MIN := 0,
       //                                                   VALUE := (SHL(IN:="AE_Position_1", N:=2) * 0.00228881) (*- "AE_Offset"*),
       //                                                   MAX := 1073741824)(*,
       //                                   MAX := "Settings_DB".VTD_Settings.VTD_Max_Heigh)*);
       // "mm_per_pulse" := 401,5584 / 262144;
       "AE_Position_1_Scaled" := (((1073741823 - (SHR(IN := "AE_Position_1", N := 2))) - 31381317) * 0.0015318237304688) - 1548572;
       // Position 2 - INPUT WORD 5 AND 6
       "AE_Position_2_Scaled" := SHR(IN := "AE_Position_2", N := 2);

       //Speed A - INPUT WORD 7
       "AE_Speed_Justified" := "AE_Speed";

       //CONTROL---------------------------------------------------------------------------------------------------------------------
       //
       //Encoder control word 2 - OUTPUT WORD 1
       //
       // 15 … 12 Master’s Sign-OF-Life (NOT relevant)
       // 10 control BY PLC 0 = No control BY the PLC 1 = Control BY the PLC Enables the PLC BY using control words TO activate / deactivate encoder functions
       // 7 Fault acknowledge Error-buffer handling NOT supported
       // 11, 9, 8, 6 … 0 Reserved
       // "AE_Control_Word_1".%X10 := "AE_PLC_Control";
       "AE_Control_Word_1".%X7 := "VTD_Reset_HMI_Tags";

       //Sensor 1 control word - OUTPUT WORD 2
       //
       // 15 Acknowledging a sensor error Description 0 = Encoder error message NOT acknowledged BY PLC 1 = Encoder error message acknowledged BY the PLC
       // 14 Activate park mode 0 = Normal operation 1 = Activate park mode
       // 13 Request FOR the absolute position value 0 = No request 1 = Request BY the master Results in the cyclic output OF the position values in G1_XIST2
       // 12 Activate preset value (see note below) Defines that a configured preset value is used (see section 3.5 on page 24) 0 = Preset value is NOT activated 1 = Preset value is activated
       // 11 Preset mode Defines how a configured preset value is used 0 = Preset value is used as a new absolute value 1 = Preset value is added TO the previous value
       // 10 … 0 Reserved
       // "AE_Control_Word_2".%X15 := "VTD_Reset_HMI_Tags";
       // "AE_Control_Word_2".%X14 := "AE_Activate_ParkMode";
       // "AE_Control_Word_2".%X13 := "AE_Request_ABS_Value";
       // "AE_Control_Word_2".%X12 := "AE_Activate_Preset_Value";
       // "AE_Control_Word_2".%X11 := "AE_Preset_Mode";
   END_REGION

   REGION LINEAR ENCODER
       "LE_X_Unsafe_Position_1" := DINT_TO_REAL("LE_X_Unsafe_Position") / 10;
       "LE_Speed_1" := "LE_Speed" * 10;
       //STATUS 
       //
       // 0 ERR - Error message (Error code in XP00– XP15); remaining bits = 0, see Error Codes
       // 1 NP - No position information/OUT (XP = 0, YP = 0, SP = 0)
       // 2 WRN - Warnings present, see Warning Module
       // 3 EV - Event present
       // 4 posdetected - Valid position information available

       //WARNINGS
       //
       // 0 WRN01 A code with non-PXV content was found.
       // 1 WRN02 the read head is too close TO the Data Matrix code tape.
       // 2 WRN03 the read head is too far from the Data Matrix code tape.
       // 3 WRN04 Y position too large. The sensor is just before OUT.
       // 4 WRN05 Y position is too small. The sensor is just before OUT.
       // 5 WRN06 the read head is rotated OR tilted in relation TO the Data Matrix code tape.
       // 6 WRN07 Low level OF code contrast.
       // 7 WRN08 Repair tape detected.
       // 8 WRN09 Temperature too high.
       // 9...15 Reserved

       //QUALITY GRADE
       //
       //The quality grades enable constant monitoring of the code tape and the camera along the entire
       //traverse distance. This enables you to detect and act upon potential damage or contamination
       //of the code tape and camera at the earliest stage possible during commissioning and normal
       //operation. As a result, this maximizes the overall functional reliability of your plant, and
       //it means you are able to immediately localize the issue in the case of a fault. Evaluations
       //are made using a scale of 1 to 6. The value 1 is the best possible read quality. A value greater
       //than 3 or worse requires the camera and its path to be inspected. The value 7 signifies "No position"
       //because no code was detected. An evaluation that indicates poor quality as the outcome can be due to
       //a misalignment or incorrect orientation, an incorrect measuring distance, or because the code tape has been affixed incorrectly
   END_REGION

       //RESET SAFETY POSITION LINEAR ENCODER
       "R_TRIG_DB_10"(CLK:="LE_Safe_Status" = 0);
       "Reintegration" := "R_TRIG_DB_10".Q;
END_FUNCTION

FUNCTION_BLOCK "FB_SICK_AFx60_PN"   // FB30, SCL
TITLE = SICK AFx60 PN
{ S7_Optimized_Access := 'TRUE' }
AUTHOR : SICKAG
FAMILY : SICKAG
VERSION : 1.1
// This function block simplifies the usage of the AFx60 encoder on Siemens S7-1200 /S7-1500 PLCs.
// It's support you to exchange the acyclic service data between the PLC and the AFx60 via Profinet (according to PROFIdrive V4.1).
// stored: AutoNumber true, IsIECCheckEnabled false, IsRetainMemResEnabled false, MemoryReserve 100, SetENOAutomatically false, UDAEnableTagReadback false
   VAR_INPUT
      ID : HW_IO;   // Hardware identifier of the "Parameter access point" module
      TOut : Time := T#5s;   // Timeout time
      Req : Bool;   // Positive trigger starts a request with the parameter set in the parameter selection
      RW : Bool;   // False= Read parameter | True= Write parameter
   END_VAR
   VAR_OUTPUT
      Done : Bool;   // The rising edge indicates if the FB processing is completed
      Busy : Bool;   // Request in process
      Error : Bool;   // Error detected
      Errorcode : "ST_SICK_AFx60_Error";   // Error code (see documentation)
   END_VAR
   VAR_IN_OUT
      Data : "ST_SICK_AFx60";   // Parameter values and data selection
   END_VAR
   VAR
      bTriggerReq { ExternalAccessible := 'False'; ExternalVisible := 'False'; ExternalWritable := 'False'} : Bool;   // Positive edge of the "Req" flag
      bTriggerReqMem { ExternalAccessible := 'False'; ExternalVisible := 'False'; ExternalWritable := 'False'} : Bool;   // Edge detection memory flag
      bTriggerReadDone { ExternalAccessible := 'False'; ExternalVisible := 'False'; ExternalWritable := 'False'} : Bool;   // Positive edge of the "RDREC.VALID" flag
      bTriggerReadDoneMem { ExternalAccessible := 'False'; ExternalVisible := 'False'; ExternalWritable := 'False'} : Bool;   // Edge detection memory flag
      bTriggerReadError { ExternalAccessible := 'False'; ExternalVisible := 'False'; ExternalWritable := 'False'} : Bool;   // Positive edge of the "RDREC.ERROR" flag
      bTriggerReadErrorMem { ExternalAccessible := 'False'; ExternalVisible := 'False'; ExternalWritable := 'False'} : Bool;   // Edge detection memory flag
      bTriggerWriteDone { ExternalAccessible := 'False'; ExternalVisible := 'False'; ExternalWritable := 'False'} : Bool;   // Positive edge of the "WRREC.DONE" flag
      bTriggerWriteDoneMem { ExternalAccessible := 'False'; ExternalVisible := 'False'; ExternalWritable := 'False'} : Bool;   // Edge detection memory flag
      bTriggerWriteError { ExternalAccessible := 'False'; ExternalVisible := 'False'; ExternalWritable := 'False'} : Bool;   // Positive edge of the "WRREC.ERROR" flag
      bTriggerWriteErrorMem { ExternalAccessible := 'False'; ExternalVisible := 'False'; ExternalWritable := 'False'} : Bool;   // Edge detection memory flag
      bRWMem { ExternalAccessible := 'False'; ExternalVisible := 'False'; ExternalWritable := 'False'} : Bool;   // Backup of the RW flag
      bBusyMem { ExternalAccessible := 'False'; ExternalVisible := 'False'; ExternalWritable := 'False'} : Bool;   // Backup of the Busy output
      iStep { ExternalAccessible := 'False'; ExternalVisible := 'False'; ExternalWritable := 'False'} : USInt;   // Program step
      iReqReference { ExternalAccessible := 'False'; ExternalVisible := 'False'; ExternalWritable := 'False'} : USInt;   // Request reference (PROFIdrive)
      iIndex { ExternalAccessible := 'False'; ExternalVisible := 'False'; ExternalWritable := 'False'} : Int;   // Temporarily variable
      iCommandIndex { ExternalAccessible := 'False'; ExternalVisible := 'False'; ExternalWritable := 'False'} : Int;   // Current command index
      fbTimeout { ExternalAccessible := 'False'; ExternalVisible := 'False'; ExternalWritable := 'False'; S7_SetPoint := 'True'} : TON_TIME;   // Instance TON
      fbReadRec { ExternalAccessible := 'False'; ExternalVisible := 'False'; ExternalWritable := 'False'; S7_SetPoint := 'True'} : RDREC;   // Instance RDREC
      fbWriteRec { ExternalAccessible := 'False'; ExternalVisible := 'False'; ExternalWritable := 'False'; S7_SetPoint := 'True'} : WRREC;   // Instance WRREC
      stTempErrorCode { ExternalAccessible := 'False'; ExternalVisible := 'False'; ExternalWritable := 'False'; S7_SetPoint := 'True'} : "ST_SICK_AFx60_Error";   // Temporariliy error code
      stRead { ExternalAccessible := 'False'; ExternalVisible := 'False'; ExternalWritable := 'False'} : Struct   // RDREC parameter
         bDone { ExternalAccessible := 'False'; ExternalVisible := 'False'; ExternalWritable := 'False'} : Bool;
         bBusy { ExternalAccessible := 'False'; ExternalVisible := 'False'; ExternalWritable := 'False'} : Bool;
         bError { ExternalAccessible := 'False'; ExternalVisible := 'False'; ExternalWritable := 'False'} : Bool;
         nStatus { ExternalAccessible := 'False'; ExternalVisible := 'False'; ExternalWritable := 'False'} : DWord;
      END_STRUCT;
      stWrite { ExternalAccessible := 'False'; ExternalVisible := 'False'; ExternalWritable := 'False'} : Struct   // WRREC parameter
         bDone { ExternalAccessible := 'False'; ExternalVisible := 'False'; ExternalWritable := 'False'} : Bool;
         bBusy { ExternalAccessible := 'False'; ExternalVisible := 'False'; ExternalWritable := 'False'} : Bool;
         bError { ExternalAccessible := 'False'; ExternalVisible := 'False'; ExternalWritable := 'False'} : Bool;
         nStatus { ExternalAccessible := 'False'; ExternalVisible := 'False'; ExternalWritable := 'False'} : DWord;
      END_STRUCT;
      arrCommandQueue { ExternalAccessible := 'False'; ExternalVisible := 'False'; ExternalWritable := 'False'} : Array[0..31] of Struct   // Command queue
         iPNU { ExternalAccessible := 'False'; ExternalVisible := 'False'; ExternalWritable := 'False'} : UInt;   // PNU
         nFormat { ExternalAccessible := 'False'; ExternalVisible := 'False'; ExternalWritable := 'False'} : Byte;   // Format
         iNoElements { ExternalAccessible := 'False'; ExternalVisible := 'False'; ExternalWritable := 'False'} : USInt;   // No. of elements
         iNoValues { ExternalAccessible := 'False'; ExternalVisible := 'False'; ExternalWritable := 'False'} : USInt;   // No. of values
      END_STRUCT;
      arrSelection { ExternalAccessible := 'False'; ExternalVisible := 'False'; ExternalWritable := 'False'} : Array[0..31] of Bool;   // Backup of the bit selection flags
      arrRecord : Array[0..254] of Byte;   // Raw data array
   END_VAR
   VAR_TEMP
      iTemp : Int;   // Temporarily variable
   END_VAR
BEGIN
   (*=============================================================================================
   Name: FB_SICK_AFx60_PN
   Author: SICK AG
   Supported PLC: S7-1200/S7-1500

   ===============================================================================================
   Description:
   This function block simplifies the usage of the AFx60 encoder on Siemens S7-1200 /S7-1500 PLCs.
   It's support you to exchange the acyclic service data between the PLC and the AFx60 via
   Profinet (according to PROFIdrive V4.1).

   The function block uses the data structure ST_SICK_AFx60 to handle data. This data structure
   includes all service data parameters of the encoder which can exchanged via the PLC.

   ===============================================================================================
   Version history:
   - - - - - - - - - - - - - - - - - - - - - - - - - - - - - - - - - - - - - - - - - - - - - - - -
   Date       | Version | Created Under        | Author  | Remark
   - - - - - - - - - - - - - - - - - - - - - - - - - - - - - - - - - - - - - - - - - - - - - - - -
   28/04/2016 | 1.0     | TIA V12 SP1 Update 4 | SICK AG | Initial version
   08/03/2017 | 1.1     | TIA V12 SP1          | SICK AG | Change units of the parameters 1002.1 
                                                           / 1003.1 from [min] to [s]

   =============================================================================================*)

   (*===================================== INITIALIZATION ======================================*)
   (*Rising edge detection*)
   #bTriggerReq:= #Req AND NOT #bTriggerReqMem;
   #bTriggerReqMem:= #Req;
   #bTriggerReadDone:= #stRead.bDone AND NOT #bTriggerReadDoneMem;
   #bTriggerReadDoneMem:= #stRead.bDone;
   #bTriggerReadError:= #stRead.bError AND NOT #bTriggerReadErrorMem;
   #bTriggerReadErrorMem:= #stRead.bError;
   #bTriggerWriteDone:= #stWrite.bDone AND NOT #bTriggerWriteDoneMem;
   #bTriggerWriteDoneMem:= #stWrite.bDone;
   #bTriggerWriteError:= #stWrite.bError AND NOT #bTriggerWriteErrorMem;
   #bTriggerWriteErrorMem:= #stWrite.bError;

   (*====================================== RECEIVE DATA =======================================*)
   #fbReadRec(ID:= #ID,
              INDEX:=16#B02E,
              MLEN:= 255,
              VALID => #stRead.bDone,
              BUSY => #stRead.bBusy,
              ERROR => #stRead.bError,
              STATUS => #stRead.nStatus,
              RECORD:= #arrRecord);
   #fbReadRec.REQ:= false;


   (*======================================== SEND DATA ========================================*)
   #fbWriteRec(ID:= #ID,
               INDEX:=16#B02E,
               DONE => #stWrite.bDone,
               BUSY => #stWrite.bBusy,
               ERROR => #stWrite.bError,
               STATUS => #stWrite.nStatus,
               RECORD:= #arrRecord);
   #fbWriteRec.REQ:= false;


   (*===================================== ERROR HANDLING ======================================*)
   IF (#stTempErrorCode.nBlockError <>0) OR (#stTempErrorCode.nCommunicationError <>0) OR (#stTempErrorCode.nEncoderError <>0) THEN
     #Done:= false;
     #Busy:= false;
     #bBusyMem:= false;
     #Error:= true;
     #Errorcode:= #stTempErrorCode;
     #stTempErrorCode.nBlockError:= 16#0000;
     #stTempErrorCode.nEncoderError:= 16#0000;
     #stTempErrorCode.nCommunicationError:= 16#0000_0000;
     #iStep:= 0;
     RETURN;
   END_IF;

   (*Time out detection*)
   #fbTimeout(IN:= #bBusyMem, PT:= #TOut);
   IF #fbTimeout.Q THEN
     #stTempErrorCode.nBlockError:= 16#0001; (*Error: Time out*)
     RETURN;
   END_IF;

   (*Read error*)
   IF #stRead.bError AND #bBusyMem THEN
     #stTempErrorCode.nBlockError:= 16#0010; (*Error: Communication error (RDREC)*)
     #stTempErrorCode.nCommunicationError:= #stRead.nStatus;
     RETURN;
   END_IF;

   (*Write error*)
   IF #stWrite.bError AND #bBusyMem THEN
     #stTempErrorCode.nBlockError:= 16#0011; (*Error: Communication error (WRREC)*)
     #stTempErrorCode.nCommunicationError:= #stWrite.nStatus;
     RETURN;
   END_IF;


   (*================================== START REQUEST (STEP 1) ==================================*)
   IF NOT #bBusyMem AND #bTriggerReq THEN
     #Done:= false;
     #Busy:= true;
     #bBusyMem:= true;
     #Error:= false;
     #Errorcode.nBlockError:= 16#0000;
     #Errorcode.nEncoderError:= 16#0000;
     #Errorcode.nCommunicationError:= 16#0000_0000;
     #bRWMem:= #RW;

     (*Save the current bit selection*)
     #arrSelection[0]:= #Data.ParameterSelection.Telegram_Number;
     #arrSelection[1]:= #Data.ParameterSelection.Device_Identification;
     #arrSelection[2]:= #Data.ParameterSelection.Enc_Profile_Number;
     #arrSelection[3]:= #Data.ParameterSelection.Eeprom_Storage;
     #arrSelection[4]:= #Data.ParameterSelection.Object_Identification;
     #arrSelection[5]:= #Data.ParameterSelection.Sensor_Format;
     #arrSelection[6]:= #Data.ParameterSelection.Parameter_List;
     #arrSelection[7]:= #Data.ParameterSelection.Encoder_Status_Flag;
     #arrSelection[8]:= #Data.ParameterSelection.Device_Status_Flag;
     #arrSelection[9]:= #Data.ParameterSelection.Diag_History_Absolute;
     #arrSelection[10]:= #Data.ParameterSelection.Diag_History_Relative;
     #arrSelection[11]:= #Data.ParameterSelection.Diag_Hist_Err_Counter;
     #arrSelection[12]:= #Data.ParameterSelection.Speed_Calculation;
     #arrSelection[13]:= #Data.ParameterSelection.Temperature_Limits;
     #arrSelection[14]:= #Data.ParameterSelection.Voltage_Limits;
     #arrSelection[15]:= #Data.ParameterSelection.Scaling_Parameters;
     #arrSelection[16]:= #Data.ParameterSelection.Operation_Test_1;
     #arrSelection[17]:= #Data.ParameterSelection.MAC_ID_Port_1;
     #arrSelection[18]:= #Data.ParameterSelection.MAC_ID_Port_2;
     #arrSelection[19]:= #Data.ParameterSelection.Version_FW_FPGA;
     #arrSelection[20]:= #Data.ParameterSelection.Temperature;
     #arrSelection[21]:= #Data.ParameterSelection.Station_Name;
     #arrSelection[22]:= #Data.ParameterSelection.Station_IP;
     #arrSelection[23]:= #Data.ParameterSelection.Station_MAC_ID;
     #arrSelection[24]:= #Data.ParameterSelection.Station_Gateway;
     #arrSelection[25]:= #Data.ParameterSelection.Station_Subnet;
     #arrSelection[26]:= #Data.ParameterSelection.Preset_Value;
     #arrSelection[27]:= #Data.ParameterSelection.Operating_Status;
     #arrSelection[28]:= false;
     #arrSelection[29]:= false;
     #arrSelection[30]:= false;
     #arrSelection[31]:= false;

     #iStep:= 2; (*Check parameter input options*)
     RETURN;
   END_IF;


   (*========================= CHECK PARAMETER INPUT OPTIONS (STEP 2) =========================*)
   IF #iStep = 2 THEN
   (*Check bit sum of the command selection*)
     #iTemp:= 0;
     FOR #iIndex:= 0 TO 31 DO
       IF #arrSelection[#iIndex] THEN
         #iTemp:= #iTemp + 1;
       END_IF;
     END_FOR;
     IF #iTemp =0 THEN
       #stTempErrorCode.nBlockError:= 16#0003; (*Error: No parameter selected (Read/Write)*)
     ELSIF #iTemp > 1 AND #bRWMem THEN
       #stTempErrorCode.nBlockError:= 16#0004; (*Error: More than one parameter selected (Write)*)
     ELSE
       #iStep:= 3; (*Creating command queue*)
     END_IF;
   END_IF;


   (*============================ CREATING COMMAND QUEUE (STEP 3) =============================*)
   IF #iStep = 3 THEN
     (*Clear command queue*)
     FOR #iIndex:= 0 TO 31 DO
       #arrCommandQueue[#iIndex].iPNU:= 0;
     END_FOR;
     #iIndex:= 0;
     #iCommandIndex:= 0;

     (*eTelegramNumber*)
     IF #arrSelection[0] THEN
       IF #bRWMem THEN
         #stTempErrorCode.nBlockError:= 16#0009; (*Error: Parameter not writable*)
       ELSE
         #arrCommandQueue[#iIndex].iPNU:= 922;
         #arrCommandQueue[#iIndex].nFormat:= 16#42;
         #arrCommandQueue[#iIndex].iNoElements:= 0;
         #arrCommandQueue[#iIndex].iNoValues:= 1;
       END_IF;
       #iIndex:= #iIndex + 1;
     END_IF;

     (*eDeviceIdentification*)
     IF #arrSelection[1] THEN
       IF #bRWMem THEN
         #stTempErrorCode.nBlockError:= 16#0009; (*Error: Parameter not writable*)
       ELSE
         #arrCommandQueue[#iIndex].iPNU:= 964;
         #arrCommandQueue[#iIndex].nFormat:= 16#42;
         #arrCommandQueue[#iIndex].iNoElements:= 6;
         #arrCommandQueue[#iIndex].iNoValues:= 6;
       END_IF;
       #iIndex:= #iIndex + 1;
     END_IF;

     (*eEncProfileNumber*)
     IF #arrSelection[2] THEN
       IF #bRWMem THEN
         #stTempErrorCode.nBlockError:= 16#0009; (*Error: Parameter not writable*)
       ELSE
         #arrCommandQueue[#iIndex].iPNU:= 965;
         #arrCommandQueue[#iIndex].nFormat:= 16#0A;
         #arrCommandQueue[#iIndex].iNoElements:= 0;
         #arrCommandQueue[#iIndex].iNoValues:= 2;
       END_IF;
       #iIndex:= #iIndex + 1;
     END_IF;

     (*eEepromStorage*)
     IF #arrSelection[3] THEN
       #arrCommandQueue[#iIndex].iPNU:= 971;
       #arrCommandQueue[#iIndex].nFormat:= 16#42;
       #arrCommandQueue[#iIndex].iNoElements:= 0;
       #arrCommandQueue[#iIndex].iNoValues:= 1;
       #iIndex:= #iIndex + 1;
     END_IF;

     (*eObjectIdentification*)
     IF #arrSelection[4] THEN
       IF #bRWMem THEN
         #stTempErrorCode.nBlockError:= 16#0009; (*Error: Parameter not writable*)
       ELSE
         #arrCommandQueue[#iIndex].iPNU:= 975;
         #arrCommandQueue[#iIndex].nFormat:= 16#42;
         #arrCommandQueue[#iIndex].iNoElements:= 7;
         #arrCommandQueue[#iIndex].iNoValues:= 7;
       END_IF;
       #iIndex:= #iIndex + 1;
     END_IF;

     (*eSensorFormat*)
     IF #arrSelection[5] THEN
       IF #bRWMem THEN
         #stTempErrorCode.nBlockError:= 16#0009; (*Error: Parameter not writable*)
       ELSE
         #arrCommandQueue[#iIndex].iPNU:= 979;
         #arrCommandQueue[#iIndex].nFormat:= 16#43;
         #arrCommandQueue[#iIndex].iNoElements:= 6;
         #arrCommandQueue[#iIndex].iNoValues:= 6;
       END_IF;
       #iIndex:= #iIndex + 1;
     END_IF;  

     (*eParameterList*)
     IF #arrSelection[6] THEN
       IF #bRWMem THEN
         #stTempErrorCode.nBlockError:= 16#0009; (*Error: Parameter not writable*)
       ELSE
         #arrCommandQueue[#iIndex].iPNU:= 980;
         #arrCommandQueue[#iIndex].nFormat:= 16#42;
         #arrCommandQueue[#iIndex].iNoElements:= 27;
         #arrCommandQueue[#iIndex].iNoValues:= 27;
       END_IF;
       #iIndex:= #iIndex + 1;
     END_IF; 

     (*eEncoderStatusFlag*)
     IF #arrSelection[7] THEN
       IF #bRWMem THEN
         #stTempErrorCode.nBlockError:= 16#0009; (*Error: Parameter not writable*)
       ELSE
         #arrCommandQueue[#iIndex].iPNU:= 1000;
         #arrCommandQueue[#iIndex].nFormat:= 16#42;
         #arrCommandQueue[#iIndex].iNoElements:= 0;
         #arrCommandQueue[#iIndex].iNoValues:= 1;
       END_IF;
       #iIndex:= #iIndex + 1;
     END_IF; 

     (*eDeviceStatusFlag*)
     IF #arrSelection[8] THEN
       IF #bRWMem THEN
         #stTempErrorCode.nBlockError:= 16#0009; (*Error: Parameter not writable*)
       ELSE
         #arrCommandQueue[#iIndex].iPNU:= 1001;
         #arrCommandQueue[#iIndex].nFormat:= 16#42;
         #arrCommandQueue[#iIndex].iNoElements:= 3;
         #arrCommandQueue[#iIndex].iNoValues:= 3;
       END_IF;
       #iIndex:= #iIndex + 1;
     END_IF; 

     (*eDiagHistoryAbsolute*)
     IF #arrSelection[9] THEN
       IF #bRWMem THEN
         #stTempErrorCode.nBlockError:= 16#0009; (*Error: Parameter not writable*)
       ELSE
         #arrCommandQueue[#iIndex].iPNU:= 1002;
         #arrCommandQueue[#iIndex].nFormat:= 16#43;
         #arrCommandQueue[#iIndex].iNoElements:= 13;
         #arrCommandQueue[#iIndex].iNoValues:= 13;
       END_IF;
       #iIndex:= #iIndex + 1;
     END_IF;   

     (*eDiagHistoryRelative*)
     IF #arrSelection[10] THEN
       IF #bRWMem THEN
         #stTempErrorCode.nBlockError:= 16#0009; (*Error: Parameter not writable*)
       ELSE
         #arrCommandQueue[#iIndex].iPNU:= 1003;
         #arrCommandQueue[#iIndex].nFormat:= 16#43;
         #arrCommandQueue[#iIndex].iNoElements:= 13;
         #arrCommandQueue[#iIndex].iNoValues:= 13;
       END_IF;
       #iIndex:= #iIndex + 1;
     END_IF;    

     (*eDiagHistErrorCounter*)
     IF #arrSelection[11] THEN
       IF #bRWMem THEN
         #stTempErrorCode.nBlockError:= 16#0009; (*Error: Parameter not writable*)
       ELSE
         #arrCommandQueue[#iIndex].iPNU:= 1004;
         #arrCommandQueue[#iIndex].nFormat:= 16#42;
         #arrCommandQueue[#iIndex].iNoElements:= 16;
         #arrCommandQueue[#iIndex].iNoValues:= 16;
       END_IF;
       #iIndex:= #iIndex + 1;
     END_IF;    

     (*eSpeedCalculation*)
     IF #arrSelection[12] THEN
       IF #bRWMem THEN
         #stTempErrorCode.nBlockError:= 16#0009; (*Error: Parameter not writable*)
       ELSE
         #arrCommandQueue[#iIndex].iPNU:= 1005;
         #arrCommandQueue[#iIndex].nFormat:= 16#42;
         #arrCommandQueue[#iIndex].iNoElements:= 6;
         #arrCommandQueue[#iIndex].iNoValues:= 6;
       END_IF;
       #iIndex:= #iIndex + 1;
     END_IF;    

     (*eTemperatureLimits*)
     IF #arrSelection[13] THEN
       #arrCommandQueue[#iIndex].iPNU:= 1006;
       #arrCommandQueue[#iIndex].nFormat:= 16#42;
       #arrCommandQueue[#iIndex].iNoElements:= 2;
       #arrCommandQueue[#iIndex].iNoValues:= 2;
       #iIndex:= #iIndex + 1;
     END_IF;    

     (*eVoltagesLimits*)
     IF #arrSelection[14] THEN
       #arrCommandQueue[#iIndex].iPNU:= 1007;
       #arrCommandQueue[#iIndex].nFormat:= 16#42;
       #arrCommandQueue[#iIndex].iNoElements:= 2;
       #arrCommandQueue[#iIndex].iNoValues:= 2;
       #iIndex:= #iIndex + 1;
     END_IF;    

     (*eScalingParameters*)
     IF #arrSelection[15] THEN
       IF #bRWMem THEN
         #stTempErrorCode.nBlockError:= 16#0009; (*Error: Parameter not writable*)
       ELSE
         #arrCommandQueue[#iIndex].iPNU:= 1009;
         #arrCommandQueue[#iIndex].nFormat:= 16#43;
         #arrCommandQueue[#iIndex].iNoElements:= 11;
         #arrCommandQueue[#iIndex].iNoValues:= 11;
       END_IF;
       #iIndex:= #iIndex + 1;
     END_IF;  

     (*eOperationTest1*)
     IF #arrSelection[16] THEN
       #arrCommandQueue[#iIndex].iPNU:= 1010;
       #arrCommandQueue[#iIndex].nFormat:= 16#42;
       #arrCommandQueue[#iIndex].iNoElements:= 0;
       #arrCommandQueue[#iIndex].iNoValues:= 1;
       #iIndex:= #iIndex + 1;
     END_IF;

     (*eMACIDPort1*)
     IF #arrSelection[17] THEN
       IF #bRWMem THEN
         #stTempErrorCode.nBlockError:= 16#0009; (*Error: Parameter not writable*)
       ELSE
         #arrCommandQueue[#iIndex].iPNU:= 1011;
         #arrCommandQueue[#iIndex].nFormat:= 16#0A;
         #arrCommandQueue[#iIndex].iNoElements:= 0;
         #arrCommandQueue[#iIndex].iNoValues:= 6;
       END_IF;
       #iIndex:= #iIndex + 1;
     END_IF;  

     (*eMACIDPort2*)
     IF #arrSelection[18] THEN
       IF #bRWMem THEN
         #stTempErrorCode.nBlockError:= 16#0009; (*Error: Parameter not writable*)
       ELSE
         #arrCommandQueue[#iIndex].iPNU:= 1012;
         #arrCommandQueue[#iIndex].nFormat:= 16#0A;
         #arrCommandQueue[#iIndex].iNoElements:= 0;
         #arrCommandQueue[#iIndex].iNoValues:= 6;
       END_IF;
       #iIndex:= #iIndex + 1;
     END_IF;

     (*eVersionFWFPGA*)
     IF #arrSelection[19] THEN
       IF #bRWMem THEN
         #stTempErrorCode.nBlockError:= 16#0009; (*Error: Parameter not writable*)
       ELSE
         #arrCommandQueue[#iIndex].iPNU:= 1013;
         #arrCommandQueue[#iIndex].nFormat:= 16#43;
         #arrCommandQueue[#iIndex].iNoElements:= 0;
         #arrCommandQueue[#iIndex].iNoValues:= 1;
       END_IF;
       #iIndex:= #iIndex + 1;
     END_IF;

     (*eTemperature*)
     IF #arrSelection[20] THEN
       IF #bRWMem THEN
         #stTempErrorCode.nBlockError:= 16#0009; (*Error: Parameter not writable*)
       ELSE
         #arrCommandQueue[#iIndex].iPNU:= 1014;
         #arrCommandQueue[#iIndex].nFormat:= 16#42;
         #arrCommandQueue[#iIndex].iNoElements:= 0;
         #arrCommandQueue[#iIndex].iNoValues:= 1;
       END_IF;
       #iIndex:= #iIndex + 1;
     END_IF;

     (*eStationName*)
     IF #arrSelection[21] THEN
       IF #bRWMem THEN
         #stTempErrorCode.nBlockError:= 16#0009; (*Error: Parameter not writable*)
       ELSE
         #arrCommandQueue[#iIndex].iPNU:= 61000;
         #arrCommandQueue[#iIndex].nFormat:= 16#0A;
         #arrCommandQueue[#iIndex].iNoElements:= 0;
         #arrCommandQueue[#iIndex].iNoValues:= 240;
       END_IF;
       #iIndex:= #iIndex + 1;
     END_IF;

     (*eStationIP*)
     IF #arrSelection[22] THEN
       IF #bRWMem THEN
         #stTempErrorCode.nBlockError:= 16#0009; (*Error: Parameter not writable*)
       ELSE
         #arrCommandQueue[#iIndex].iPNU:= 61001;
         #arrCommandQueue[#iIndex].nFormat:= 16#43;
         #arrCommandQueue[#iIndex].iNoElements:= 0;
         #arrCommandQueue[#iIndex].iNoValues:= 1;
       END_IF;
       #iIndex:= #iIndex + 1;
     END_IF;

     (*eStationMACID*)
     IF #arrSelection[23] THEN
       IF #bRWMem THEN
         #stTempErrorCode.nBlockError:= 16#0009; (*Error: Parameter not writable*)
       ELSE
         #arrCommandQueue[#iIndex].iPNU:= 61002;
         #arrCommandQueue[#iIndex].nFormat:= 16#0A;
         #arrCommandQueue[#iIndex].iNoElements:= 0;
         #arrCommandQueue[#iIndex].iNoValues:= 6;
       END_IF;
       #iIndex:= #iIndex + 1;
     END_IF;

     (*eStationGateway*)
     IF #arrSelection[24] THEN
       IF #bRWMem THEN
         #stTempErrorCode.nBlockError:= 16#0009; (*Error: Parameter not writable*)
       ELSE
         #arrCommandQueue[#iIndex].iPNU:= 61003;
         #arrCommandQueue[#iIndex].nFormat:= 16#43;
         #arrCommandQueue[#iIndex].iNoElements:= 0;
         #arrCommandQueue[#iIndex].iNoValues:= 1;
       END_IF;
       #iIndex:= #iIndex + 1;
     END_IF;

     (*eStationSubnet*)
     IF #arrSelection[25] THEN
       IF #bRWMem THEN
         #stTempErrorCode.nBlockError:= 16#0009; (*Error: Parameter not writable*)
       ELSE
         #arrCommandQueue[#iIndex].iPNU:= 61004;
         #arrCommandQueue[#iIndex].nFormat:= 16#43;
         #arrCommandQueue[#iIndex].iNoElements:= 0;
         #arrCommandQueue[#iIndex].iNoValues:= 1;
       END_IF;
       #iIndex:= #iIndex + 1;
     END_IF;

     (*ePresetValue*)
     IF #arrSelection[26] THEN
       #arrCommandQueue[#iIndex].iPNU:= 65000;
       #arrCommandQueue[#iIndex].nFormat:= 16#43;
       #arrCommandQueue[#iIndex].iNoElements:= 0;
       #arrCommandQueue[#iIndex].iNoValues:= 1;
       #iIndex:= #iIndex + 1;
     END_IF;

     (*eOperatingStatus*)
     IF #arrSelection[27] THEN
       IF #bRWMem THEN
         #stTempErrorCode.nBlockError:= 16#0009; (*Error: Parameter not writable*)
       ELSE
         #arrCommandQueue[#iIndex].iPNU:= 65001;
         #arrCommandQueue[#iIndex].nFormat:= 16#43;
         #arrCommandQueue[#iIndex].iNoElements:= 12;
         #arrCommandQueue[#iIndex].iNoValues:= 12;
       END_IF;
       #iIndex:= #iIndex + 1;
     END_IF;

     (*Check if no error occurs while validation*)
     IF #stTempErrorCode.nBlockError = 0 THEN
       #iStep:= 4; (*Check communication status*)
     END_IF;
   END_IF;


   (*========================== CHECK COMMUNICATION STATUS (STEP 4) ==========================*)
   IF #iStep = 4 THEN
     IF NOT #stRead.bBusy AND NOT #stWrite.bBusy THEN
       #iStep:= 5; (*Send request*)
     END_IF;
   END_IF;


   (*================================= SEND REQUEST (STEP 5) =================================*)
   IF #iStep = 5 THEN

     (*Request reference calculation*)
     #iReqReference:= #iReqReference + 1;
     IF #iReqReference = 0 THEN
       #iReqReference:= 1;
     END_IF;

     (*Request parameter*)
     #arrRecord[0]:= #iReqReference; (*Request reference*)
     IF #bRWMem THEN
       #arrRecord[1]:= 2; (*Request ID = Change parameter*)
     ELSE
       #arrRecord[1]:= 1; (*Request ID = Request parameter*)
     END_IF;
     #arrRecord[2]:= 0; (*DO-ID*)
     #arrRecord[3]:= 1; (*No. of parameters*)
     #arrRecord[4]:= 16#10; (*Attribute = Value*)
     #arrRecord[5]:= #arrCommandQueue[#iCommandIndex].iNoElements; (*No. of elements*)
     #arrRecord[6]:= #arrCommandQueue[#iCommandIndex].iPNU.%B1; (*PNU high byte*)
     #arrRecord[7]:= #arrCommandQueue[#iCommandIndex].iPNU.%B0; (*PNU low byte*)
     #arrRecord[8]:= 0; (*Subindex high byte*)
     #arrRecord[9]:= 0; (*Subindex low byte*)
     #fbWriteRec.REQ:= true;

     (*Add parameter value*)
     IF #bRWMem THEN
       #arrRecord[10]:= #arrCommandQueue[#iCommandIndex].nFormat;
       #arrRecord[11]:= #arrCommandQueue[#iCommandIndex].iNoValues;

       CASE #arrCommandQueue[#iCommandIndex].iPNU OF
         (*eEepromStorage*)
         971:
           #arrRecord[12]:= #Data.Parameter.Eeprom_Storage.%B1;
           #arrRecord[13]:= #Data.Parameter.Eeprom_Storage.%B0;

         (*eTemperatureLimits*)
         1006:
           #arrRecord[12]:= #Data.Parameter.Temperature_Limits.Lower_Limit.%B1;
           #arrRecord[13]:= #Data.Parameter.Temperature_Limits.Lower_Limit.%B0;
           #arrRecord[14]:= #Data.Parameter.Temperature_Limits.Upper_Limit.%B1;
           #arrRecord[15]:= #Data.Parameter.Temperature_Limits.Upper_Limit.%B0;

         (*eVoltageLimits*)
         1007:
           #arrRecord[12]:= #Data.Parameter.Voltage_Limits.Lower_Limit.%B1;
           #arrRecord[13]:= #Data.Parameter.Voltage_Limits.Lower_Limit.%B0;
           #arrRecord[14]:= #Data.Parameter.Voltage_Limits.Upper_Limit.%B1;
           #arrRecord[15]:= #Data.Parameter.Voltage_Limits.Upper_Limit.%B0;

         (*eOperationTest1*)
         1010:
           #arrRecord[12]:= #Data.Parameter.Operation_Test_1.%B1;
           #arrRecord[13]:= #Data.Parameter.Operation_Test_1.%B0;

         (*ePresetValue*)
         65000:
           #arrRecord[12]:= #Data.Parameter.Preset_Value.%B3;
           #arrRecord[13]:= #Data.Parameter.Preset_Value.%B2;
           #arrRecord[14]:= #Data.Parameter.Preset_Value.%B1;
           #arrRecord[15]:= #Data.Parameter.Preset_Value.%B0;     
         ELSE
           #stTempErrorCode.nBlockError:= 16#0002; (*Error: Internal error*)
           RETURN;
         END_CASE;

       (*Add telegram length (write)*)
       IF #arrCommandQueue[#iCommandIndex].nFormat = 16#41 THEN
         #fbWriteRec.LEN:= 12 + #arrCommandQueue[#iCommandIndex].iNoValues; (*Byte*)
       ELSIF #arrCommandQueue[#iCommandIndex].nFormat = 16#42 THEN
         #fbWriteRec.LEN:= 12 + (#arrCommandQueue[#iCommandIndex].iNoValues * 2); (*Word*)
       ELSIF #arrCommandQueue[#iCommandIndex].nFormat =16#43 THEN
         #fbWriteRec.LEN:= 12 + (#arrCommandQueue[#iCommandIndex].iNoValues * 4); (*DWord*)
       ELSE
         #stTempErrorCode.nBlockError:= 16#0002; (*Error: Internal error*)
         RETURN;
       END_IF;
     ELSE
       (*Add telegram length (read)*)
       #fbWriteRec.LEN:= 10;
     END_IF;

     #iStep:= 6; (*Waiting for a write response*)
   END_IF;


   (*========================== WAITING FOR A WRITE RESPONSE (STEP 6) ==========================*)
   IF #iStep = 6 THEN
     IF #stWrite.bDone THEN
       #fbReadRec.REQ:= true;
       #iStep:= 7;
       RETURN;
     END_IF;
   END_IF;


   (*========================== WAITING FOR A READ RESPONSE (STEP 7) ===========================*)
   IF #iStep = 7 THEN
     IF #stRead.bDone THEN

       (*Check: Request reference*)
       IF #iReqReference <> #arrRecord[0] THEN
         #stTempErrorCode.nBlockError:= 16#0005; (*Error: Invalid request reference received*)
         RETURN;
       END_IF;

       (*Check: Response negative*)
       IF #arrRecord[4] = 16#44 THEN
         #stTempErrorCode.nBlockError:= 16#000A; (*Error: Encoder error*)
         #stTempErrorCode.nEncoderError.%B0:= #arrRecord[7];
         #stTempErrorCode.nEncoderError.%B1:= #arrRecord[6];
         RETURN;
       END_IF;

       (*Check: Response positive*)
       IF #arrRecord[4] = 16#40 THEN
         #iStep:= 9; (*Action permormed / Next command*)
       ELSE
         #iStep:= 8; (*Check response data*)
       END_IF;
     END_IF;
   END_IF;


   (*============================= CHECKING RESPONSE DATA (STEP 8) =============================*)
   IF #iStep = 8 THEN
     (*Check: Data type format*)
     IF #arrRecord[4] <> #arrCommandQueue[#iCommandIndex].nFormat THEN
       #stTempErrorCode.nBlockError:= 16#0006; (*Error: Unexpected data type format received*)
       RETURN;

     (*Check: No. of values*)
     ELSIF (#arrRecord[5] <> #arrCommandQueue[#iCommandIndex].iNoValues) AND (#arrRecord[4] <> 16#0A) THEN
       #stTempErrorCode.nBlockError:= 16#0007; (*Error: Unexpected no. of values received*)
       RETURN;
     END_IF;

     (*Get value*)
     CASE #arrCommandQueue[#iCommandIndex].iPNU OF
       (*eTelegramNumber*)
       922:
         #Data.Parameter.Telegram_Number.%B0:= #arrRecord[7];
         #Data.Parameter.Telegram_Number.%B1:= #arrRecord[8];

       (*eDeviceIdentification*)
       964:
         #Data.Parameter.Device_Identification.Manufacturer.%B1:= #arrRecord[6];
         #Data.Parameter.Device_Identification.Manufacturer.%B0:= #arrRecord[7];
         #Data.Parameter.Device_Identification.Encoder_Unit_Type.%B1:= #arrRecord[8];
         #Data.Parameter.Device_Identification.Encoder_Unit_Type.%B0:= #arrRecord[9];
         #Data.Parameter.Device_Identification.FW_Version.%B1:= #arrRecord[10];
         #Data.Parameter.Device_Identification.FW_Version.%B0:= #arrRecord[11];
         #Data.Parameter.Device_Identification.FW_Date_Year.%B1:= #arrRecord[12];
         #Data.Parameter.Device_Identification.FW_Date_Year.%B0:= #arrRecord[13];
         #Data.Parameter.Device_Identification.FW_Date_Day_Month.%B1:= #arrRecord[14];
         #Data.Parameter.Device_Identification.FW_Date_Day_Month.%B0:= #arrRecord[15];
         #Data.Parameter.Device_Identification.Number_Of_Objects.%B1:= #arrRecord[16];
         #Data.Parameter.Device_Identification.Number_Of_Objects.%B0:= #arrRecord[17];

       (*eEncProfileNumber*)
       965:
         #Data.Parameter.Enc_Profile_Number.Profile_Number:= #arrRecord[6];
         #Data.Parameter.Enc_Profile_Number.Profile_Version:= #arrRecord[7];

       (*eEepromStorage*)
       971:
         #Data.Parameter.Eeprom_Storage.%B1:= #arrRecord[6];
         #Data.Parameter.Eeprom_Storage.%B0:= #arrRecord[7];

       (*eObjectIdentification*)
       975:
         #Data.Parameter.Object_Identification.Manufacturer.%B1:= #arrRecord[6];
         #Data.Parameter.Object_Identification.Manufacturer.%B0:= #arrRecord[7];
         #Data.Parameter.Object_Identification.Encoder_Unit_Type.%B1:= #arrRecord[8];
         #Data.Parameter.Object_Identification.Encoder_Unit_Type.%B0:= #arrRecord[9];
         #Data.Parameter.Object_Identification.FW_Version.%B1:= #arrRecord[10];
         #Data.Parameter.Object_Identification.FW_Version.%B0:= #arrRecord[11];
         #Data.Parameter.Object_Identification.FW_Date_Year.%B1:= #arrRecord[12];
         #Data.Parameter.Object_Identification.FW_Date_Year.%B0:= #arrRecord[13];
         #Data.Parameter.Object_Identification.FW_Date_Day_Month.%B1:= #arrRecord[14];
         #Data.Parameter.Object_Identification.FW_Date_Day_Month.%B0:= #arrRecord[15];  
         #Data.Parameter.Object_Identification.EO_Type_Class.%B1:= #arrRecord[16];
         #Data.Parameter.Object_Identification.EO_Type_Class.%B0:= #arrRecord[17];
         #Data.Parameter.Object_Identification.EO_Sub_Class.%B1:= #arrRecord[18];
         #Data.Parameter.Object_Identification.EO_Sub_Class.%B0:= #arrRecord[19];

       (*eSensorFormat*)
       979:
         #Data.Parameter.Sensor_Format.Header.%B3:= #arrRecord[6];
         #Data.Parameter.Sensor_Format.Header.%B2:= #arrRecord[7];
         #Data.Parameter.Sensor_Format.Header.%B1:= #arrRecord[8];
         #Data.Parameter.Sensor_Format.Header.%B0:= #arrRecord[9];
         #Data.Parameter.Sensor_Format.Sensor_Type.%B3:= #arrRecord[10];
         #Data.Parameter.Sensor_Format.Sensor_Type.%B2:= #arrRecord[11];
         #Data.Parameter.Sensor_Format.Sensor_Type.%B1:= #arrRecord[12];
         #Data.Parameter.Sensor_Format.Sensor_Type.%B0:= #arrRecord[13];
         #Data.Parameter.Sensor_Format.Sensor_Resolution.%B3:= #arrRecord[14];
         #Data.Parameter.Sensor_Format.Sensor_Resolution.%B2:= #arrRecord[15];
         #Data.Parameter.Sensor_Format.Sensor_Resolution.%B1:= #arrRecord[16];
         #Data.Parameter.Sensor_Format.Sensor_Resolution.%B0:= #arrRecord[17];
         #Data.Parameter.Sensor_Format.Shift_Factor_Left.%B3:= #arrRecord[18];
         #Data.Parameter.Sensor_Format.Shift_Factor_Left.%B2:= #arrRecord[19];
         #Data.Parameter.Sensor_Format.Shift_Factor_Left.%B1:= #arrRecord[20];
         #Data.Parameter.Sensor_Format.Shift_Factor_Left.%B0:= #arrRecord[21];
         #Data.Parameter.Sensor_Format.Shift_Factor_Right.%B3:= #arrRecord[22];
         #Data.Parameter.Sensor_Format.Shift_Factor_Right.%B2:= #arrRecord[23];
         #Data.Parameter.Sensor_Format.Shift_Factor_Right.%B1:= #arrRecord[24];
         #Data.Parameter.Sensor_Format.Shift_Factor_Right.%B0:= #arrRecord[25];
         #Data.Parameter.Sensor_Format.Revolutions.%B3:= #arrRecord[26];
         #Data.Parameter.Sensor_Format.Revolutions.%B2:= #arrRecord[27];
         #Data.Parameter.Sensor_Format.Revolutions.%B1:= #arrRecord[28];
         #Data.Parameter.Sensor_Format.Revolutions.%B0:= #arrRecord[29];

       (*eParameterList*)
       980:
         FOR #iIndex:= 0 TO 26 DO
           #Data.Parameter.Parameter_List[#iIndex].%B1:= #arrRecord[6 + 2 * #iIndex];
           #Data.Parameter.Parameter_List[#iIndex].%B0:= #arrRecord[7 + 2 * #iIndex];
         END_FOR;

       (*eEncoderStatusFlag*)
       1000:
         #Data.Parameter.Encoder_Status_Flag.%B1:= #arrRecord[6];
         #Data.Parameter.Encoder_Status_Flag.%B0:= #arrRecord[7];

       (*eDeviceStatusFlag*)
       1001:
         #Data.Parameter.Device_Status_Flag.S_STAT_A.%B1:= #arrRecord[6];
         #Data.Parameter.Device_Status_Flag.S_STAT_A.%B0:= #arrRecord[7];
         #Data.Parameter.Device_Status_Flag.S_STAT_B.%B1:= #arrRecord[8];
         #Data.Parameter.Device_Status_Flag.S_STAT_B.%B0:= #arrRecord[9];      
         #Data.Parameter.Device_Status_Flag.S_STAT_C.%B1:= #arrRecord[10];
         #Data.Parameter.Device_Status_Flag.S_STAT_C.%B0:= #arrRecord[11];

